// TwinCAT 3 PLC project HrlRbgPlc
// ProgramVersion: 3.1.4026.25
// libraries:
//   NodeTree, * (sulemanali5760)
//   Tc2_MC2, * (Beckhoff Automation GmbH)
//   Tc3_JsonXml, * (Beckhoff Automation GmbH)
//   Tc2_TcpIp, * (Beckhoff Automation GmbH)
//   Tc2_Standard, * (Beckhoff Automation GmbH)
//   Tc2_System, * (Beckhoff Automation GmbH)
//   TcUnit, * (www.tcunit.org)
// project tree:
//   / PlcTask.TcTTO
//   Rack/ GVL_Rack.TcGVL, ST_Slot.TcDUT, ST_SlotAddr.TcDUT, FB_Rack.TcPOU
//   Devices/ E_IPointResult.TcDUT, E_ZoneState.TcDUT, E_AxisKind.TcDUT, I_Axis.TcIO, FB_AxisNc.TcPOU, FB_Axis.TcPOU, FB_ConveyorZone.TcPOU, FB_IPoint.TcPOU
//   Performance/ ST_SrmKinematics.TcDUT, F_DoubleCycleTime.TcPOU, F_LoadHandlingTime.TcPOU, F_MoveTime.TcPOU, F_TravelTime.TcPOU
//   Units/ FB_Srm.TcPOU, E_JogAxis.TcDUT
//   Mfr/ GVL_Mfr.TcGVL, ST_Telegram.TcDUT, FB_MfrInterface.TcPOU, E_MfrLink.TcDUT, ST_TelegramLayout.TcDUT, I_MfrLink.TcIO, FB_TelegramCodec.TcPOU, FB_MfrLinkTcp.TcPOU
//   Machine/ FB_Hrl.TcPOU, FB_MfrEmulator.TcPOU, MAIN.TcPOU
//   Test/ GVL_Test.TcGVL, FB_Axis_Test.TcPOU, FB_ConveyorZone_Test.TcPOU, FB_IPoint_Test.TcPOU, FB_MfrInterface_Test.TcPOU, FB_Rack_Test.TcPOU, FB_Srm_Test.TcPOU, FB_TravelTime_Test.TcPOU, FB_AxisNc_Test.TcPOU, FB_HrlConfig_Test.TcPOU, FB_MfrLinkFake.TcPOU, FB_TelegramCodec_Test.TcPOU, FB_Operation_Test.TcPOU, FB_SafetyInterface_Test.TcPOU, PRG_TEST.TcPOU
//   Config/ ST_RackConfig.TcDUT, ST_AxisConfig.TcDUT, ST_ZoneConfig.TcDUT, ST_HrlConfig.TcDUT, FB_HrlConfig.TcPOU
//   Commissioning/ FB_TeachIn.TcPOU
//   Diag/ E_Fault.TcDUT, FB_Diag.TcPOU
//   Safety/ ST_SafetyStatus.TcDUT, FB_SafetyInterface.TcPOU
//   Hmi/ ST_HmiStatus.TcDUT, ST_HmiCommand.TcDUT, GVL_Hmi.TcGVL, FB_HmiBridge.TcPOU
// real-time tasks:
//   TASK PlcTask: cycle T#10ms, priority 20, ADS port 350
// motion (NC):
//   TASK NC-Task 1 SAF: cycle T#2ms, priority 4, ADS port 501
//   TASK NC-Task 1 SVB: cycle T#10ms, priority 8, ADS port 511
//   AXIS Travel (id 1)
//     Velo: Fast=3000, Maximum=3500
//     OtherSettings: AllowMotionCmdToSlave=true
//     encoder EncType=1
//     drive DrvType=5
//       Analog: VeloReferenz=3500, TorqueSetpointScale=10, ScaleFactorActTorque=0.1
//       TimeComp: TaskDelayCycles=1
//     controller CtrType=1
//       CtrPara: PriorControlFactor=1
//         Observer: BandWidth=20
//   AXIS Hoist (id 2)
//     OtherSettings: AllowMotionCmdToSlave=true
//     encoder EncType=1
//     drive DrvType=5
//       Analog: TorqueSetpointScale=10, ScaleFactorActTorque=0.1
//       TimeComp: TaskDelayCycles=1
//     controller CtrType=1
//       CtrPara: PriorControlFactor=1
//         Observer: BandWidth=20
//   AXIS Fork (id 3)
//     OtherSettings: AllowMotionCmdToSlave=true
//     encoder EncType=1
//     drive DrvType=5
//       Analog: TorqueSetpointScale=10, ScaleFactorActTorque=0.1
//       TimeComp: TaskDelayCycles=1
//     controller CtrType=1
//       CtrPara: PriorControlFactor=1
//         Observer: BandWidth=20
//   AXIS TestAxis (id 4)
//     OtherSettings: AllowMotionCmdToSlave=true
//     encoder EncType=1
//     drive DrvType=5
//       Analog: TorqueSetpointScale=10, ScaleFactorActTorque=0.1
//       TimeComp: TaskDelayCycles=1
//     controller CtrType=1
//       CtrPara: PriorControlFactor=1
//         Observer: BandWidth=20
//   AXIS TestTravel (id 5)
//     Velo: Fast=3000, Maximum=3500
//     OtherSettings: AllowMotionCmdToSlave=true
//     encoder EncType=1
//     drive DrvType=5
//       Analog: VeloReferenz=3500, TorqueSetpointScale=10, ScaleFactorActTorque=0.1
//       TimeComp: TaskDelayCycles=1
//     controller CtrType=1
//       CtrPara: PriorControlFactor=1
//         Observer: BandWidth=20
//   AXIS TestHoist (id 6)
//     OtherSettings: AllowMotionCmdToSlave=true
//     encoder EncType=1
//     drive DrvType=5
//       Analog: TorqueSetpointScale=10, ScaleFactorActTorque=0.1
//       TimeComp: TaskDelayCycles=1
//     controller CtrType=1
//       CtrPara: PriorControlFactor=1
//         Observer: BandWidth=20
//   AXIS TestFork (id 7)
//     OtherSettings: AllowMotionCmdToSlave=true
//     encoder EncType=1
//     drive DrvType=5
//       Analog: TorqueSetpointScale=10, ScaleFactorActTorque=0.1
//       TimeComp: TaskDelayCycles=1
//     controller CtrType=1
//       CtrPara: PriorControlFactor=1
//         Observer: BandWidth=20
// variable links:
//   HrlRbgPlc/HrlRbgPlc Instance <-> NC-Task 1 SAF/Axes/Fork
//     PlcTask Inputs/MAIN.fbPlant.fbSrm.fbForkNc.stAxis.NcToPlc <-> Outputs/ToPlc
//     PlcTask Outputs/MAIN.fbPlant.fbSrm.fbForkNc.stAxis.PlcToNc <-> Inputs/FromPlc
//   HrlRbgPlc/HrlRbgPlc Instance <-> NC-Task 1 SAF/Axes/Hoist
//     PlcTask Inputs/MAIN.fbPlant.fbSrm.fbHoistNc.stAxis.NcToPlc <-> Outputs/ToPlc
//     PlcTask Outputs/MAIN.fbPlant.fbSrm.fbHoistNc.stAxis.PlcToNc <-> Inputs/FromPlc
//   HrlRbgPlc/HrlRbgPlc Instance <-> NC-Task 1 SAF/Axes/TestAxis
//     PlcTask Inputs/PRG_TEST.fbAxisNcTest.fbAxis.stAxis.NcToPlc <-> Outputs/ToPlc
//     PlcTask Outputs/PRG_TEST.fbAxisNcTest.fbAxis.stAxis.PlcToNc <-> Inputs/FromPlc
//   HrlRbgPlc/HrlRbgPlc Instance <-> NC-Task 1 SAF/Axes/TestFork
//     PlcTask Inputs/PRG_TEST.fbAxisNcTest.fbSrmNc.fbForkNc.stAxis.NcToPlc <-> Outputs/ToPlc
//     PlcTask Outputs/PRG_TEST.fbAxisNcTest.fbSrmNc.fbForkNc.stAxis.PlcToNc <-> Inputs/FromPlc
//   HrlRbgPlc/HrlRbgPlc Instance <-> NC-Task 1 SAF/Axes/TestHoist
//     PlcTask Inputs/PRG_TEST.fbAxisNcTest.fbSrmNc.fbHoistNc.stAxis.NcToPlc <-> Outputs/ToPlc
//     PlcTask Outputs/PRG_TEST.fbAxisNcTest.fbSrmNc.fbHoistNc.stAxis.PlcToNc <-> Inputs/FromPlc
//   HrlRbgPlc/HrlRbgPlc Instance <-> NC-Task 1 SAF/Axes/TestTravel
//     PlcTask Inputs/PRG_TEST.fbAxisNcTest.fbSrmNc.fbTravelNc.stAxis.NcToPlc <-> Outputs/ToPlc
//     PlcTask Outputs/PRG_TEST.fbAxisNcTest.fbSrmNc.fbTravelNc.stAxis.PlcToNc <-> Inputs/FromPlc
//   HrlRbgPlc/HrlRbgPlc Instance <-> NC-Task 1 SAF/Axes/Travel
//     PlcTask Inputs/MAIN.fbPlant.fbSrm.fbTravelNc.stAxis.NcToPlc <-> Outputs/ToPlc
//     PlcTask Outputs/MAIN.fbPlant.fbSrm.fbTravelNc.stAxis.PlcToNc <-> Inputs/FromPlc

CONFIGURATION HrlRbgPlc
    RESOURCE PLC ON TwinCAT3
        TASK PlcTask(INTERVAL := T#10ms, PRIORITY := 20);
        PROGRAM MAIN WITH PlcTask : MAIN;
        PROGRAM PRG_TEST WITH PlcTask : PRG_TEST;
    END_RESOURCE
END_CONFIGURATION

// ---- Rack/ST_Slot.TcDUT
TYPE ST_Slot :
STRUCT
    bOccupied : BOOL;
    sLeId     : STRING(20);   // load unit id (pallet barcode)
    bTaught   : BOOL;         // TRUE once the place was measured in teach mode
    lrTaughtX : LREAL;        // measured travel position [m]
    lrTaughtY : LREAL;        // measured hoist position [m]
END_STRUCT
END_TYPE

// ---- Rack/ST_SlotAddr.TcDUT
// Address of a storage place, as the material flow computer sends it.
// Column 0 / level 1 / side 1 is the transfer station (Uebergabeplatz) at the
// front of the aisle, where the pre-zone hands pallets to the RBG.
TYPE ST_SlotAddr :
STRUCT
    nSide   : INT;   // 1 = left, 2 = right (seen from the transfer station)
    nColumn : INT;   // 1..GVL_Rack.cColumns, 0 = transfer station
    nLevel  : INT;   // 1..GVL_Rack.cLevels
END_STRUCT
END_TYPE

// ---- Devices/E_IPointResult.TcDUT
{attribute 'qualified_only'}
{attribute 'strict'}
TYPE E_IPointResult :
(
    eOk         := 0,   // contour fine, barcode read -> may be stored
    eNioContour := 1,   // overhang or too high -> back to the operator
    eNioNoRead  := 2    // barcode not readable -> back to the operator
) DINT;
END_TYPE

// ---- Devices/E_ZoneState.TcDUT
{attribute 'qualified_only'}
{attribute 'strict'}
TYPE E_ZoneState :
(
    eEmpty      := 0,
    eReceiving  := 1,   // motor on, pallet running in
    eOccupied   := 2,   // pallet at the end light barrier, motor off
    eDelivering := 3,   // motor on, pallet running out to the next zone
    eFault      := 4    // jam (light barrier not reached in time) or drive fault
) DINT;
END_TYPE

// ---- Devices/E_AxisKind.TcDUT
// Which implementation drives the RBG axes. Switched in the configuration,
// never in the code: the sequence only talks to I_Axis.
{attribute 'qualified_only'}
{attribute 'strict'}
TYPE E_AxisKind :
(
    eSim := 0,   // FB_Axis: simulated trapezoid profile, simulated time (tests, demo)
    eNc  := 1    // FB_AxisNc: Beckhoff NC axis via Tc2_MC2 (real drive or NC simulation axis)
) INT;
END_TYPE

// ---- Performance/ST_SrmKinematics.TcDUT
TYPE ST_SrmKinematics :
STRUCT
    lrVeloX  : LREAL;   // travel
    lrAccelX : LREAL;
    lrVeloY  : LREAL;   // hoist
    lrAccelY : LREAL;
    lrVeloZ  : LREAL;   // telescopic fork
    lrAccelZ : LREAL;
END_STRUCT
END_TYPE

// ---- Mfr/ST_Telegram.TcDUT
// One telegram between the material flow computer (MFR, e.g. WAMAS) and the PLC.
// The real WAMAS layout is project-specific; this is a typical fixed layout.
TYPE ST_Telegram :
STRUCT
    sType    : STRING(4);    // TORD order, TACK acknowledge, TDON done, TERR error
    nSeq     : UINT;         // sequence number of the sender, +1 per telegram
    nOrder   : DINT;         // transport order number
    sLeId    : STRING(20);   // load unit id
    stSource : ST_SlotAddr;
    stTarget : ST_SlotAddr;
    nStatus  : INT;          // GVL_Mfr status codes, 0 = OK
END_STRUCT
END_TYPE

// ---- Config/ST_RackConfig.TcDUT
// Rack geometry of one aisle. Defaults = the practice plant (GVL_Rack).
// Sizes may not exceed GVL_Rack.cMaxSides / cMaxColumns / cMaxLevels.
TYPE ST_RackConfig :
STRUCT
    nSides          : INT   := GVL_Rack.cSides;
    nColumns        : INT   := GVL_Rack.cColumns;
    nLevels         : INT   := GVL_Rack.cLevels;
    lrPitchX        : LREAL := GVL_Rack.cPitchX;          // column pitch incl. upright [m]
    lrPitchY        : LREAL := GVL_Rack.cPitchY;          // level pitch [m]
    lrOffsetX       : LREAL := GVL_Rack.cOffsetX;         // transfer station -> centre of column 1 [m]
    lrOffsetY       : LREAL := GVL_Rack.cOffsetY;         // fork height at level 1 / station [m]
    lrForkStroke    : LREAL := GVL_Rack.cForkStroke;      // [m]
    lrLiftStroke    : LREAL := GVL_Rack.cLiftStroke;      // [m]
    lrTeachTolerance: LREAL := GVL_Rack.cTeachTolerance;  // [m]
END_STRUCT
END_TYPE

// ---- Config/ST_AxisConfig.TcDUT
TYPE ST_AxisConfig :
STRUCT
    lrVelocity : LREAL := 1.0;   // [m/s]
    lrAccel    : LREAL := 0.5;   // acceleration = deceleration [m/s2]
END_STRUCT
END_TYPE

// ---- Config/ST_ZoneConfig.TcDUT
// Parameters of one conveyor zone (the standard block FB_ConveyorZone).
TYPE ST_ZoneConfig :
STRUCT
    lrLength     : LREAL := 1.6;    // up to the end light barrier [m]
    lrSpeed      : LREAL := 0.2;    // [m/s]
    lrJamTimeout : LREAL := 20.0;   // [s]
    bSimulate    : BOOL  := TRUE;   // FALSE: end light barrier from the real input
END_STRUCT
END_TYPE

// ---- Config/ST_HrlConfig.TcDUT
// Everything an integrator sets per plant. Loaded from HrlConfig.json by
// FB_HrlConfig; every default here is the practice plant, so a missing file
// or a missing entry still gives a working demo.
TYPE ST_HrlConfig :
STRUCT
    stRack    : ST_RackConfig;
    eAxisKind : E_AxisKind := E_AxisKind.eSim;
    stTravel  : ST_AxisConfig := (lrVelocity := 3.0, lrAccel := 0.6);
    stHoist   : ST_AxisConfig := (lrVelocity := 1.5, lrAccel := 0.8);
    stFork    : ST_AxisConfig := (lrVelocity := 0.6, lrAccel := 0.6);
    stInfeed  : ST_ZoneConfig;
    stOutfeed : ST_ZoneConfig := (lrLength := 2.4, lrSpeed := 0.2, lrJamTimeout := 20.0, bSimulate := TRUE);
    lrAckTimeout : LREAL := 5.0;   // MFR must acknowledge TDON within this [s]
    eMfrLink     : E_MfrLink := E_MfrLink.eEmulator;
    nMfrPort     : UINT := 2000;    // TCP port the PLC listens on (eTcp)
    stLayout     : ST_TelegramLayout;
    bSafetySimulate : BOOL := TRUE;   // bench without safety controller (never on a real machine)
END_STRUCT
END_TYPE

// ---- Mfr/E_MfrLink.TcDUT
// Where the transport orders come from.
{attribute 'qualified_only'}
{attribute 'strict'}
TYPE E_MfrLink :
(
    eEmulator := 0,   // FB_MfrEmulator in the PLC (commissioning, demo, tests)
    eTcp      := 1    // real material flow computer over TCP/IP (PLC is the server)
) INT;
END_TYPE

// ---- Mfr/ST_TelegramLayout.TcDUT
// Field widths of the fixed-length ASCII telegram. The field order is fixed:
//   type | seq | order | load unit | source side,column,level | target side,column,level | status
// Numbers are right-aligned with leading zeros, the load unit id is
// left-aligned and padded with spaces. The frame is STX + fields + ETX.
// Defaults give a 52-character telegram.
TYPE ST_TelegramLayout :
STRUCT
    nType   : INT := 4;
    nSeq    : INT := 5;
    nOrder  : INT := 8;
    nLeId   : INT := 20;
    nSide   : INT := 1;
    nColumn : INT := 3;
    nLevel  : INT := 2;
    nStatus : INT := 3;
END_STRUCT
END_TYPE

// ---- Units/E_JogAxis.TcDUT
// Axis the operator jogs in manual mode.
{attribute 'qualified_only'}
{attribute 'strict'}
TYPE E_JogAxis :
(
    eTravel := 0,
    eHoist  := 1,
    eFork   := 2
) INT;
END_TYPE

// ---- Diag/E_Fault.TcDUT
// Plant faults reported by FB_Diag (index into its active list).
{attribute 'qualified_only'}
{attribute 'strict'}
TYPE E_Fault :
(
    eSrmAxis      := 1,   // an RBG axis failed during a job
    eInfeedJam    := 2,
    eOutfeedJam   := 3,
    eMfrAck       := 4,   // MFR did not acknowledge TDON in time
    eMfrLinkDown  := 5,   // TCP link configured but no MFR connected
    eConfig       := 6,   // HrlConfig.json rejected, defaults in use
    eTeachRejected:= 7,   // measured place too far from the drawing
    eSafety       := 8    // safety stop or restart lock active
) INT;
END_TYPE

// ---- Safety/ST_SafetyStatus.TcDUT
// Status bits the safety controller (e.g. TwinSAFE logic) gives the standard
// PLC. The standard PLC only reads them: it never switches safety itself.
// Map each bit to the TwinSAFE group output (see docs/safety/README.md).
TYPE ST_SafetyStatus :
STRUCT
    bSafetyRun  : BOOL;   // safety program running, no group error
    bEStopOk    : BOOL;   // all emergency stops released
    bDoorClosed : BOOL;   // aisle access door closed
    bDoorLocked : BOOL;   // aisle access door guard-locked
    bStoOk      : BOOL;   // drives not in Safe Torque Off
END_STRUCT
END_TYPE

// ---- Hmi/ST_HmiStatus.TcDUT
// Everything the HMI shows (PLC -> HMI). Filled by MAIN every cycle.
TYPE ST_HmiStatus :
STRUCT
    nMode          : INT;          // 0 stop, 1 manual, 2 homing, 3 automatic (E_OpMode)
    bSafetyOk      : BOOL;
    lrTravelPos    : LREAL;        // [m]
    lrHoistPos     : LREAL;        // [m]
    lrForkPos      : LREAL;        // [m]
    bBusy          : BOOL;         // RBG job running
    bFault         : BOOL;         // RBG fault, needs reset
    bJogBlocked    : BOOL;         // jog refused: fork not centred
    sLeOnFork      : STRING(20);
    nJobsDone      : DINT;
    nStored        : DINT;         // emulator counters
    nRetrieved     : DINT;
    bMfrConnected  : BOOL;         // TCP link (always FALSE with the emulator)
    nActiveFaults  : INT;
    sFault1        : STRING(80);   // first four active faults, cause - remedy
    sFault2        : STRING(80);
    sFault3        : STRING(80);
    sFault4        : STRING(80);
    bTeachActive   : BOOL;
    nTaught        : INT;
    bTeachRejected : BOOL;
    sConfigError   : STRING(120);
END_STRUCT
END_TYPE

// ---- Hmi/ST_HmiCommand.TcDUT
// Everything the HMI may command (HMI -> PLC). Buttons that trigger an action
// (teach start/confirm, resets) are evaluated on the rising edge in MAIN.
TYPE ST_HmiCommand :
STRUCT
    bModeStop     : BOOL;       // mode buttons: TRUE while pressed (button state symbol)
    bModeManual   : BOOL;
    bModeHoming   : BOOL;
    bModeAuto     : BOOL;
    nJogAxis      : INT;        // 0 travel, 1 hoist, 2 fork
    bJogFwd       : BOOL;       // held while the button is pressed
    bJogBwd       : BOOL;
    nTeachSide    : INT := 1;
    nTeachColumn  : INT := 1;
    nTeachLevel   : INT := 1;
    bTeachStart   : BOOL;
    bTeachConfirm : BOOL;
    bResetFault   : BOOL;       // RBG fault reset
    bSafetyReset  : BOOL;       // safety acknowledge
END_STRUCT
END_TYPE

// ---- Rack/GVL_Rack.TcGVL
{attribute 'qualified_only'}
VAR_GLOBAL CONSTANT
    // Largest rack the PLC reserves memory for. The real size comes from the
    // configuration (ST_RackConfig) and may be anything up to these.
    cMaxSides   : INT   := 2;
    cMaxColumns : INT   := 60;
    cMaxLevels  : INT   := 16;
    // Defaults = the practice plant: one aisle, single-deep, both sides.
    cSides      : INT   := 2;
    cColumns    : INT   := 20;
    cLevels     : INT   := 8;
    cPitchX     : LREAL := 1.40;   // column pitch incl. upright [m]
    cPitchY     : LREAL := 1.30;   // level pitch [m]
    cOffsetX    : LREAL := 2.00;   // transfer station -> centre of column 1 [m]
    cOffsetY    : LREAL := 0.50;   // fork height at level 1 / transfer station [m]
    cForkStroke : LREAL := 1.10;   // telescopic fork travel into a place [m]
    cLiftStroke : LREAL := 0.10;   // lift to take a pallet off its beams [m]
    // Teach-in: a measured place may differ from the drawing by this much;
    // more means a bent or wrongly built rack -> reject and check the rack.
    cTeachTolerance : LREAL := 0.020;   // [m]
END_VAR

// ---- Mfr/GVL_Mfr.TcGVL
{attribute 'qualified_only'}
VAR_GLOBAL CONSTANT
    cStatusOk         : INT := 0;
    cSlotOccupied     : INT := 10;   // target place occupied
    cSlotEmpty        : INT := 11;   // source place empty
    cContourNio       : INT := 20;   // pallet failed the I-point
    cAckTimeout       : INT := 30;   // MFR did not acknowledge TDON in time
    cWrongSequence    : INT := 40;   // telegram sequence number out of order
    cDuplicateOrder   : INT := 41;   // order number already active / just done
    cInvalidAddress   : INT := 42;
    cSrmBusy          : INT := 43;
    cLeMismatch       : INT := 44;   // load unit at the source is not the one ordered
    cUnknownTelegram  : INT := 45;
    cSrmFault         : INT := 50;
END_VAR

// ---- Test/GVL_Test.TcGVL
{attribute 'qualified_only'}
VAR_GLOBAL
    // Results of the FEM 9.851 double-cycle test, for the performance protocol.
    lrDoubleCycleCalc     : LREAL;   // calculated [s]
    lrDoubleCycleMeasured : LREAL;   // measured in the simulation [s]
    lrDoubleCyclesPerHour : LREAL;   // 3600 / measured
END_VAR

// ---- Hmi/GVL_Hmi.TcGVL
// The only PLC data the HMI uses. Both structs are mapped automatically into
// the TwinCAT HMI server (attribute TcHmiSymbol.AddSymbol).
{attribute 'qualified_only'}
VAR_GLOBAL
    {attribute 'TcHmiSymbol.AddSymbol'}
    stStatus  : ST_HmiStatus;
    {attribute 'TcHmiSymbol.AddSymbol'}
    stCommand : ST_HmiCommand;
END_VAR

// ---- Devices/I_Axis.TcIO
// I_Axis - what the RBG sequence needs from a positioning axis, whatever
// drives it: the simulated FB_Axis or the NC axis FB_AxisNc. Units are metres.
INTERFACE I_Axis

// Drive to an absolute position: eBusy while moving, eDone in position, eError on a fault.
METHOD MoveAbs : E_CmdResult
VAR_INPUT
    lrPos : LREAL;   // target [m]
END_VAR
END_METHOD

// Acknowledge a fault: the axis stops where it is and waits for a new target.
METHOD Reset
VAR_INPUT
END_VAR
END_METHOD

// Stop now (end of a jog, stop mode). The axis then waits for a new target.
METHOD Halt
VAR_INPUT
END_VAR
END_METHOD

// Actual position [m].
PROPERTY ActPos : LREAL
GET
END_GET
END_PROPERTY

PROPERTY Error : BOOL
GET
END_GET
END_PROPERTY

END_INTERFACE

// ---- Mfr/I_MfrLink.TcIO
// I_MfrLink - transport of telegrams between the PLC and the material flow
// computer. FB_MfrInterface only sees telegrams; how they travel (TCP, a test
// double) is behind this interface.
INTERFACE I_MfrLink

// Next received telegram, TRUE if there was one. A frame that could not be
// decoded comes back with sType = 'BAD'.
METHOD Poll : BOOL
VAR_IN_OUT
    stIn : ST_Telegram;
END_VAR
END_METHOD

// Queue a telegram for the MFR. FALSE if not connected or the queue is full.
METHOD Send : BOOL
VAR_INPUT
    stOut : ST_Telegram;
END_VAR
END_METHOD

PROPERTY Connected : BOOL
GET
END_GET
END_PROPERTY

END_INTERFACE

// ---- Machine/MAIN.TcPOU
// MAIN - builds the plant from HrlConfig.json, runs it in the operating mode
// the HMI asks for (eModeRequest), forced to stop while the safety interface
// does not allow motion. With mfr.link = emulator the MFR emulator drives it.
// Watch fbPlant.fbSrm (positions, jobs), fbPlant.fbRack and fbPlant.fbDiag online.
PROGRAM MAIN
VAR
    fbPlant      : FB_Hrl(ipParent := 0, sNodeName := 'HRL');
    fbOpMode     : FB_OpModeHandler;
    fbEmulator   : FB_MfrEmulator;
    fbConfig     : FB_HrlConfig;   // HrlConfig.json from the boot folder; defaults if absent
    fbHmi        : FB_HmiBridge;   // GVL_Hmi <-> plant
    eModeNow     : E_OpMode;
    bInit        : BOOL := TRUE;
END_VAR

IF bInit THEN
    fbConfig();
    IF NOT fbConfig.bDone THEN
        RETURN;   // the plant starts only with its final configuration
    END_IF
    fbPlant.stConfig     := fbConfig.stConfig;
    fbPlant.sConfigError := fbConfig.sError;
    fbOpMode.SetRoot(fbPlant);
    bInit := FALSE;
END_IF

fbHmi.Run(fbPlant, fbEmulator, GVL_Hmi.stCommand, GVL_Hmi.stStatus, eModeNow);
IF fbPlant.bSafetyOk THEN
    eModeNow := fbHmi.eModeRequest;
ELSE
    eModeNow := E_OpMode.eStop;   // safety first: no motion without the safety OK
END_IF
fbOpMode.Mode := eModeNow;
IF fbPlant.stConfig.eMfrLink = E_MfrLink.eEmulator THEN
    fbEmulator.Run(fbPlant);   // no real MFR: the emulator sends the orders
END_IF
fbOpMode.Cyclic();

END_PROGRAM

// ---- Machine/FB_Hrl.TcPOU
// FB_Hrl - the whole practice plant as the root mode node: one aisle with one
// RBG, the rack, the pre-zone with I-point and in-feed/out-feed conveyors, and
// the MFR interface.
// Pre-zone flow: in-feed (pallet already checked at the I-point) -> transfer
// station -> RBG stores it. Retrieved pallets are put on the station and leave
// over the out-feed.
FUNCTION_BLOCK FB_Hrl EXTENDS FB_ModeNode
VAR_INPUT
    stConfig : ST_HrlConfig;   // applied once on the first cycle (set it before)
    sConfigError : STRING(120);   // from FB_HrlConfig; shown as a fault
    stSafety     : ST_SafetyStatus;   // map from the safety controller (TwinSAFE group outputs)
    bSafetyReset : BOOL;              // acknowledge button
    bDoorRequest : BOOL;              // operator wants to enter the aisle
END_VAR
VAR
    fbRack    : FB_Rack;
    fbSrm     : FB_Srm(ipParent := THIS^, sNodeName := 'RBG01');
    fbInfeed  : FB_ConveyorZone(ipParent := THIS^, sNodeName := 'Infeed');
    fbOutfeed : FB_ConveyorZone(ipParent := THIS^, sNodeName := 'Outfeed');
    fbIPoint  : FB_IPoint;
    fbMfr     : FB_MfrInterface;
    fbMfrTcp  : FB_MfrLinkTcp;     // used when stConfig.eMfrLink = eTcp
    fbTeach   : FB_TeachIn;        // guided teach-in (manual mode)
    fbDiag    : FB_Diag;           // active faults for the HMI + TwinCAT logger
    fbSafety  : FB_SafetyInterface;
    bInitDone : BOOL;
    nInStep   : INT;
    sMovingLe : STRING(20);
END_VAR
VAR_OUTPUT
    bStationOutbound : BOOL;   // pallet on the station is leaving (retrieved), not arriving
    bStationReserved : BOOL;   // station held free for a retrieval: the in-feed must wait
    bSafetyOk        : BOOL;   // drives may run; FALSE -> MAIN forces stop mode
    bDoorUnlockReq   : BOOL;   // to the safety controller
END_VAR

METHOD PROTECTED OnCyclic
VAR_INPUT
END_VAR
IF NOT bInitDone THEN
    // The plant is built from the configuration; the code below never changes per site.
    fbRack.stCfg      := stConfig.stRack;
    fbSrm.eAxisKind   := stConfig.eAxisKind;
    fbSrm.stTravelCfg := stConfig.stTravel;
    fbSrm.stHoistCfg  := stConfig.stHoist;
    fbSrm.stForkCfg   := stConfig.stFork;
    ApplyZone(fbInfeed, stConfig.stInfeed);    // same standard block, other parameters
    ApplyZone(fbOutfeed, stConfig.stOutfeed);
    fbMfr.lrAckTimeout := stConfig.lrAckTimeout;
    fbSrm.Init(fbRack);
    fbMfr.Init(fbRack, fbSrm);
    fbTeach.Init(fbRack, fbSrm);
    fbMfrTcp.nPort    := stConfig.nMfrPort;
    fbMfrTcp.stLayout := stConfig.stLayout;
    bInitDone := TRUE;
END_IF
IF stConfig.eMfrLink = E_MfrLink.eTcp THEN
    fbMfrTcp.Cyclic();          // the link stays up in every operating mode
    fbMfr.Serve(fbMfrTcp);
END_IF
fbSafety(stStatus := stSafety, bSimulate := stConfig.bSafetySimulate, bReset := bSafetyReset,
         bDoorRequest := bDoorRequest, bStandstill := NOT fbSrm.bBusy AND NOT fbSrm.bGotoActive);
bSafetyOk      := fbSafety.bDriveEnable;
bDoorUnlockReq := fbSafety.bDoorUnlockReq;
SUPER^.OnCyclic();
fbDiag.Check(E_Fault.eSafety, NOT bSafetyOk, 'Safety stop - check e-stop and aisle door, then acknowledge');
fbDiag.Check(E_Fault.eSrmAxis, fbSrm.bFault, 'RBG axis fault - check the drive, then ResetFault');
fbDiag.Check(E_Fault.eInfeedJam, fbInfeed.eState = E_ZoneState.eFault, 'In-feed jam - clear the pallet, reset the zone');
fbDiag.Check(E_Fault.eOutfeedJam, fbOutfeed.eState = E_ZoneState.eFault, 'Out-feed jam - clear the pallet, reset the zone');
fbDiag.Check(E_Fault.eMfrAck, fbMfr.bAckTimeout, 'MFR did not acknowledge TDON - check the MFR');
fbDiag.Check(E_Fault.eMfrLinkDown, stConfig.eMfrLink = E_MfrLink.eTcp AND NOT fbMfrTcp.bConnected,
             'No MFR connected - check network / MFR port');
fbDiag.Check(E_Fault.eConfig, sConfigError <> '', 'HrlConfig.json rejected - defaults in use, see sConfigError');
fbDiag.Check(E_Fault.eTeachRejected, fbTeach.bLastRejected, 'Teach-in refused - place too far from drawing, check rack');
END_METHOD

METHOD PROTECTED RunAutomatic
VAR_INPUT
END_VAR
VAR
    stStation : ST_SlotAddr := (nSide := 1, nColumn := 0, nLevel := 1);
END_VAR
fbMfr.Cyclic();

// In-feed -> transfer station
CASE nInStep OF
    0:  IF fbInfeed.eState = E_ZoneState.eOccupied AND NOT fbRack.IsOccupied(stStation)
           AND NOT bStationOutbound AND NOT bStationReserved THEN
            sMovingLe := fbInfeed.sLeId;
            nInStep   := 1;
        END_IF
    // Done once our pallet has left the zone. The previous zone may hand over
    // the next pallet in the same cycle, so "zone empty" alone can be missed.
    1:  IF fbInfeed.Deliver() = E_CmdResult.eDone OR fbInfeed.sLeId <> sMovingLe THEN
            fbRack.Put(stStation, sMovingLe);
            nInStep := 0;
        END_IF
END_CASE

// Transfer station -> out-feed (only pallets the RBG brought out)
IF bStationOutbound AND fbRack.IsOccupied(stStation)
   AND fbOutfeed.eState = E_ZoneState.eEmpty THEN
    fbOutfeed.Accept(fbRack.Take(stStation));
    bStationOutbound := FALSE;
    bStationReserved := FALSE;   // station free for the in-feed again
END_IF
IF fbOutfeed.eState = E_ZoneState.eOccupied THEN
    fbOutfeed.Deliver();   // goods-out takes it away
END_IF
END_METHOD

// Called when a retrieval to the station is ordered: that pallet leaves.
METHOD PUBLIC MarkStationOutbound
VAR_INPUT
END_VAR
bStationOutbound := TRUE;
END_METHOD

// Hold the transfer station free for the next retrieval. Without this the
// in-feed refills the station every time the RBG picks a pallet from it, and
// a retrieval never finds the station empty.
METHOD PUBLIC ReserveStation
VAR_INPUT
END_VAR
bStationReserved := TRUE;
END_METHOD

// Manual jog request from the HMI (acts in manual mode only).
METHOD PUBLIC Jog
VAR_INPUT
    eAxis : E_JogAxis;
    bFwd  : BOOL;
    bBwd  : BOOL;
END_VAR
fbSrm.eJogAxis := eAxis;
fbSrm.bJogFwd  := bFwd;
fbSrm.bJogBwd  := bBwd;
END_METHOD

METHOD PRIVATE ApplyZone
VAR_IN_OUT
    fbZone : FB_ConveyorZone;
END_VAR
VAR_INPUT
    stCfg : ST_ZoneConfig;
END_VAR
fbZone.lrLength     := stCfg.lrLength;
fbZone.lrSpeed      := stCfg.lrSpeed;
fbZone.lrJamTimeout := stCfg.lrJamTimeout;
fbZone.bSimulate    := stCfg.bSimulate;
END_METHOD

END_FUNCTION_BLOCK

// ---- Rack/FB_Rack.TcPOU
// FB_Rack - the PLC's picture of the rack: which place is occupied by which
// load unit, and where each place really is (nominal from the drawing, or the
// value measured during teach-in). It is data, not a machine node, so the RBG,
// the MFR interface and the tests all share one instance by reference.
FUNCTION_BLOCK FB_Rack
VAR_INPUT
    stCfg : ST_RackConfig;   // geometry; set once before the first job (FB_Hrl does it from the config)
END_VAR
VAR
    aSlot     : ARRAY[1..GVL_Rack.cMaxSides, 1..GVL_Rack.cMaxColumns, 1..GVL_Rack.cMaxLevels] OF ST_Slot;
    stStation : ST_Slot;   // the transfer station in front of the aisle
END_VAR

METHOD PUBLIC IsStation : BOOL
VAR_INPUT
    stAddr : ST_SlotAddr;
END_VAR
IsStation := stAddr.nColumn = 0 AND stAddr.nLevel = 1 AND stAddr.nSide = 1;
END_METHOD

METHOD PUBLIC IsValid : BOOL
VAR_INPUT
    stAddr : ST_SlotAddr;
END_VAR
IsValid := IsStation(stAddr)
        OR (stAddr.nSide >= 1 AND stAddr.nSide <= stCfg.nSides
            AND stAddr.nColumn >= 1 AND stAddr.nColumn <= stCfg.nColumns
            AND stAddr.nLevel >= 1 AND stAddr.nLevel <= stCfg.nLevels);
END_METHOD

// Pointer to the place record, or 0 for an invalid address.
METHOD PRIVATE Slot : POINTER TO ST_Slot
VAR_INPUT
    stAddr : ST_SlotAddr;
END_VAR
IF IsStation(stAddr) THEN
    Slot := ADR(stStation);
ELSIF IsValid(stAddr) THEN
    Slot := ADR(aSlot[stAddr.nSide, stAddr.nColumn, stAddr.nLevel]);
ELSE
    Slot := 0;
END_IF
END_METHOD

// Travel position of a place from the drawing [m].
METHOD PUBLIC NominalX : LREAL
VAR_INPUT
    stAddr : ST_SlotAddr;
END_VAR
IF IsStation(stAddr) THEN
    NominalX := 0.0;
ELSE
    NominalX := stCfg.lrOffsetX + INT_TO_LREAL(stAddr.nColumn - 1) * stCfg.lrPitchX;
END_IF
END_METHOD

// Hoist position of a place from the drawing [m].
METHOD PUBLIC NominalY : LREAL
VAR_INPUT
    stAddr : ST_SlotAddr;
END_VAR
NominalY := stCfg.lrOffsetY + INT_TO_LREAL(stAddr.nLevel - 1) * stCfg.lrPitchY;
END_METHOD

// Where the RBG drives to: the taught position if there is one, else nominal.
METHOD PUBLIC TargetX : LREAL
VAR_INPUT
    stAddr : ST_SlotAddr;
END_VAR
VAR
    pSlot : POINTER TO ST_Slot;
END_VAR
pSlot := Slot(stAddr);
IF pSlot <> 0 AND_THEN pSlot^.bTaught THEN
    TargetX := pSlot^.lrTaughtX;
ELSE
    TargetX := NominalX(stAddr);
END_IF
END_METHOD

METHOD PUBLIC TargetY : LREAL
VAR_INPUT
    stAddr : ST_SlotAddr;
END_VAR
VAR
    pSlot : POINTER TO ST_Slot;
END_VAR
pSlot := Slot(stAddr);
IF pSlot <> 0 AND_THEN pSlot^.bTaught THEN
    TargetY := pSlot^.lrTaughtY;
ELSE
    TargetY := NominalY(stAddr);
END_IF
END_METHOD

// Store the measured position of a place (teach-in). Returns FALSE and keeps
// the old value if the measurement is further than cTeachTolerance from the
// drawing - that is a rack to check, not a value to learn.
METHOD PUBLIC Teach : BOOL
VAR_INPUT
    stAddr : ST_SlotAddr;
    lrX    : LREAL;   // measured travel position [m] (laser distance sensor)
    lrY    : LREAL;   // measured hoist position [m]
END_VAR
VAR
    pSlot : POINTER TO ST_Slot;
END_VAR
pSlot := Slot(stAddr);
IF pSlot = 0 OR IsStation(stAddr)
   OR ABS(lrX - NominalX(stAddr)) > stCfg.lrTeachTolerance
   OR ABS(lrY - NominalY(stAddr)) > stCfg.lrTeachTolerance THEN
    Teach := FALSE;
    RETURN;
END_IF
pSlot^.lrTaughtX := lrX;
pSlot^.lrTaughtY := lrY;
pSlot^.bTaught   := TRUE;
Teach := TRUE;
END_METHOD

METHOD PUBLIC IsOccupied : BOOL
VAR_INPUT
    stAddr : ST_SlotAddr;
END_VAR
VAR
    pSlot : POINTER TO ST_Slot;
END_VAR
pSlot := Slot(stAddr);
IsOccupied := pSlot <> 0 AND_THEN pSlot^.bOccupied;
END_METHOD

METHOD PUBLIC LeIdAt : STRING(20)
VAR_INPUT
    stAddr : ST_SlotAddr;
END_VAR
VAR
    pSlot : POINTER TO ST_Slot;
END_VAR
pSlot := Slot(stAddr);
IF pSlot <> 0 AND_THEN pSlot^.bOccupied THEN
    LeIdAt := pSlot^.sLeId;
ELSE
    LeIdAt := '';
END_IF
END_METHOD

// Book a load unit into a place. FALSE if the place is invalid or occupied.
METHOD PUBLIC Put : BOOL
VAR_INPUT
    stAddr : ST_SlotAddr;
    sLeId  : STRING(20);
END_VAR
VAR
    pSlot : POINTER TO ST_Slot;
END_VAR
pSlot := Slot(stAddr);
IF pSlot = 0 OR_ELSE pSlot^.bOccupied OR sLeId = '' THEN
    Put := FALSE;
    RETURN;
END_IF
pSlot^.bOccupied := TRUE;
pSlot^.sLeId     := sLeId;
Put := TRUE;
END_METHOD

// Book a load unit out of a place; returns its id, or '' if the place was empty.
METHOD PUBLIC Take : STRING(20)
VAR_INPUT
    stAddr : ST_SlotAddr;
END_VAR
VAR
    pSlot : POINTER TO ST_Slot;
END_VAR
pSlot := Slot(stAddr);
IF pSlot = 0 OR_ELSE NOT pSlot^.bOccupied THEN
    Take := '';
    RETURN;
END_IF
Take := pSlot^.sLeId;
pSlot^.bOccupied := FALSE;
pSlot^.sLeId     := '';
END_METHOD

// First free place, filled column by column from the transfer station
// (short travel first). FALSE if the rack is full.
METHOD PUBLIC FindFree : BOOL
VAR_IN_OUT
    stFound : ST_SlotAddr;
END_VAR
VAR
    nCol, nLvl, nSide : INT;
END_VAR
FOR nCol := 1 TO stCfg.nColumns DO
    FOR nLvl := 1 TO stCfg.nLevels DO
        FOR nSide := 1 TO stCfg.nSides DO
            IF NOT aSlot[nSide, nCol, nLvl].bOccupied THEN
                stFound.nSide   := nSide;
                stFound.nColumn := nCol;
                stFound.nLevel  := nLvl;
                FindFree := TRUE;
                RETURN;
            END_IF
        END_FOR
    END_FOR
END_FOR
FindFree := FALSE;
END_METHOD

END_FUNCTION_BLOCK

// ---- Units/FB_Srm.TcPOU
// FB_Srm - the storage and retrieval machine (Regalbediengeraet, RBG) as a
// mode node. Its three axes are child device nodes, so one Cyclic() on the RBG
// runs the sequence first and then lets the axes move in the same scan.
//
// A job moves one load unit from a source place to a target place (either may
// be the transfer station). The sequence is the classic single cycle:
//   travel+hoist to source -> fork out -> lift -> fork in ->
//   travel+hoist to target (loaded, lifted) -> fork out -> lower -> fork in.
// Two jobs back to back (store, then retrieve) make a double cycle.
FUNCTION_BLOCK FB_Srm EXTENDS FB_ModeNode
VAR_INPUT
    eAxisKind : E_AxisKind := E_AxisKind.eSim;   // simulated axes or NC axes
    stTravelCfg : ST_AxisConfig := (lrVelocity := 3.0, lrAccel := 0.6);
    stHoistCfg  : ST_AxisConfig := (lrVelocity := 1.5, lrAccel := 0.8);
    stForkCfg   : ST_AxisConfig := (lrVelocity := 0.6, lrAccel := 0.6);
    // Manual mode (HMI): hold bJogFwd / bJogBwd to move eJogAxis, release to stop.
    eJogAxis : E_JogAxis := E_JogAxis.eTravel;
    bJogFwd  : BOOL;
    bJogBwd  : BOOL;
END_VAR
VAR_OUTPUT
    bBusy         : BOOL;         // a job is running
    bJobDone      : BOOL;         // last job finished; stays TRUE until the next StartJob
    bFault        : BOOL;         // sequence stopped on an axis fault -> ResetFault
    nJobsDone     : DINT;
    lrLastJobTime : LREAL;        // simulated duration of the last job [s]
    sLeOnFork     : STRING(20);   // load unit currently on the fork
    bJogBlocked   : BOOL;         // jog refused: fork not centred for travel / hoist
    bGotoActive   : BOOL;         // manual: driving to a GotoXY target (teach-in)
END_VAR
VAR
    fbTravel : FB_Axis(ipParent := THIS^, sNodeName := 'Travel');
    fbHoist  : FB_Axis(ipParent := THIS^, sNodeName := 'Hoist');
    fbFork   : FB_Axis(ipParent := THIS^, sNodeName := 'Fork');
    fbTravelNc : FB_AxisNc(ipParent := THIS^, sNodeName := 'TravelNc');
    fbHoistNc  : FB_AxisNc(ipParent := THIS^, sNodeName := 'HoistNc');
    fbForkNc   : FB_AxisNc(ipParent := THIS^, sNodeName := 'ForkNc');
    ipTravel : I_Axis;   // the axes the sequence uses, chosen by eAxisKind
    ipHoist  : I_Axis;
    ipFork   : I_Axis;
    fbCycle  : FB_CycleManager;
    refRack  : REFERENCE TO FB_Rack;
    stSource : ST_SlotAddr;
    stTarget : ST_SlotAddr;
    bJobPending : BOOL;
    lrJobTime   : LREAL;
    lrGotoX     : LREAL;
    lrGotoY     : LREAL;
    bJogging    : BOOL;
END_VAR

// Give the RBG the rack it works on (once, before the first job).
METHOD PUBLIC Init
VAR_INPUT
    fbRackRef : REFERENCE TO FB_Rack;
END_VAR
refRack REF= fbRackRef;
END_METHOD

// Accept a transport job. FALSE if busy, faulted, the addresses are invalid,
// the source is empty or the target is occupied.
METHOD PUBLIC StartJob : BOOL
VAR_INPUT
    stFrom : ST_SlotAddr;
    stTo   : ST_SlotAddr;
END_VAR
StartJob := FALSE;
IF NOT __ISVALIDREF(refRack) OR bJobPending OR bFault THEN
    RETURN;
END_IF
IF NOT refRack.IsValid(stFrom) OR NOT refRack.IsValid(stTo)
   OR NOT refRack.IsOccupied(stFrom) OR refRack.IsOccupied(stTo) THEN
    RETURN;
END_IF
stSource    := stFrom;
stTarget    := stTo;
lrJobTime   := 0.0;
bJobDone    := FALSE;
bJobPending := TRUE;
fbCycle.Reset();   // so the next Call() sees a fresh start edge
StartJob := TRUE;
END_METHOD

// Acknowledge a fault. A load unit still on the fork stays booked on the fork.
METHOD PUBLIC ResetFault
VAR_INPUT
END_VAR
SelectAxes();
ipTravel.Reset();
ipHoist.Reset();
ipFork.Reset();
fbCycle.Reset();
bFault      := FALSE;
bJobPending := FALSE;
END_METHOD

// Travel and hoist together; done when both are in position.
METHOD PRIVATE MoveXY : E_CmdResult
VAR_INPUT
    lrX : LREAL;
    lrY : LREAL;
END_VAR
VAR
    eX, eY : E_CmdResult;
END_VAR
eX := ipTravel.MoveAbs(lrX);
eY := ipHoist.MoveAbs(lrY);
IF eX = E_CmdResult.eError OR eY = E_CmdResult.eError THEN
    MoveXY := E_CmdResult.eError;
ELSIF eX = E_CmdResult.eDone AND eY = E_CmdResult.eDone THEN
    MoveXY := E_CmdResult.eDone;
ELSE
    MoveXY := E_CmdResult.eBusy;
END_IF
END_METHOD

// Fork end position for a place: left side (and the station) negative, right positive.
METHOD PRIVATE ForkPos : LREAL
VAR_INPUT
    stAddr : ST_SlotAddr;
END_VAR
IF stAddr.nSide = 2 THEN
    ForkPos := refRack.stCfg.lrForkStroke;
ELSE
    ForkPos := -refRack.stCfg.lrForkStroke;
END_IF
END_METHOD

METHOD PROTECTED OnCyclic
VAR_INPUT
END_VAR
SelectAxes();
// Axis data from the configuration (defaults = the practice RBG).
fbTravel.lrVelocity   := stTravelCfg.lrVelocity;  fbTravel.lrAccel   := stTravelCfg.lrAccel;
fbHoist.lrVelocity    := stHoistCfg.lrVelocity;   fbHoist.lrAccel    := stHoistCfg.lrAccel;
fbFork.lrVelocity     := stForkCfg.lrVelocity;    fbFork.lrAccel     := stForkCfg.lrAccel;
fbTravelNc.lrVelocity := stTravelCfg.lrVelocity;  fbTravelNc.lrAccel := stTravelCfg.lrAccel;
fbHoistNc.lrVelocity  := stHoistCfg.lrVelocity;   fbHoistNc.lrAccel  := stHoistCfg.lrAccel;
fbForkNc.lrVelocity   := stForkCfg.lrVelocity;    fbForkNc.lrAccel   := stForkCfg.lrAccel;
IF bJobPending THEN
    lrJobTime := lrJobTime + fbTravel.lrCycleTime;
END_IF
SUPER^.OnCyclic();   // dispatch to RunAutomatic / RunManual / ...
bBusy := bJobPending;
END_METHOD

METHOD PROTECTED RunAutomatic
VAR_INPUT
END_VAR
IF NOT __ISVALIDREF(refRack) THEN
    RETURN;
END_IF

fbCycle.Call(bExecute := bJobPending);
CASE fbCycle.Step OF
    0:  fbCycle.Await(MoveXY(refRack.TargetX(stSource), refRack.TargetY(stSource)));
    1:  fbCycle.Await(ipFork.MoveAbs(ForkPos(stSource)));
    2:  IF fbCycle.Await(ipHoist.MoveAbs(refRack.TargetY(stSource) + refRack.stCfg.lrLiftStroke)) THEN
            sLeOnFork := refRack.Take(stSource);   // pallet is now on the fork
        END_IF
    3:  fbCycle.Await(ipFork.MoveAbs(0.0));
    4:  fbCycle.Await(MoveXY(refRack.TargetX(stTarget), refRack.TargetY(stTarget) + refRack.stCfg.lrLiftStroke));
    5:  fbCycle.Await(ipFork.MoveAbs(ForkPos(stTarget)));
    6:  IF fbCycle.Await(ipHoist.MoveAbs(refRack.TargetY(stTarget))) THEN
            refRack.Put(stTarget, sLeOnFork);      // pallet is on the beams
            sLeOnFork := '';
        END_IF
    7:  IF fbCycle.Await(ipFork.MoveAbs(0.0)) THEN
            bJobPending   := FALSE;
            bJobDone      := TRUE;
            nJobsDone     := nJobsDone + 1;
            lrLastJobTime := lrJobTime;
        END_IF
END_CASE

IF fbCycle.Error THEN
    bFault := TRUE;
END_IF
END_METHOD

// Go to the transfer station: fork in first, then travel and hoist.
METHOD PROTECTED RunHoming
VAR_INPUT
END_VAR
IF NOT __ISVALIDREF(refRack) THEN
    RETURN;
END_IF
IF ipFork.MoveAbs(0.0) = E_CmdResult.eDone THEN
    MoveXY(0.0, refRack.stCfg.lrOffsetY);
END_IF
END_METHOD

PROPERTY PUBLIC TravelPos : LREAL
GET
SelectAxes();
TravelPos := ipTravel.ActPos;
END_GET
END_PROPERTY

PROPERTY PUBLIC HoistPos : LREAL
GET
SelectAxes();
HoistPos := ipHoist.ActPos;
END_GET
END_PROPERTY

PROPERTY PUBLIC ForkActPos : LREAL
GET
SelectAxes();
ForkActPos := ipFork.ActPos;
END_GET
END_PROPERTY

// Test and commissioning aid: simulate a fault of the travel drive.
METHOD PUBLIC InjectTravelFault
VAR_INPUT
    bFaultOn : BOOL;
END_VAR
fbTravel.bDriveFault := bFaultOn;
END_METHOD

// Manual mode: drive travel and hoist to a position (fork stays centred).
// Used by teach-in to go to the nominal position of a place.
METHOD PUBLIC GotoXY : BOOL
VAR_INPUT
    lrX : LREAL;
    lrY : LREAL;
END_VAR
IF bFault OR bJobPending THEN
    RETURN;
END_IF
lrGotoX     := lrX;
lrGotoY     := lrY;
bGotoActive := TRUE;
GotoXY      := TRUE;
END_METHOD

// Jog one axis while a button is held; travel and hoist only with the fork
// centred (a fork in the rack would hit the uprights). A GotoXY target has
// priority over jogging.
METHOD PROTECTED RunManual
VAR_INPUT
END_VAR
VAR
    ipAx    : I_Axis;
    lrLimit : LREAL;
END_VAR
IF NOT __ISVALIDREF(refRack) THEN
    RETURN;
END_IF
IF bGotoActive THEN
    IF ABS(ipFork.ActPos) > 0.005 THEN
        ipFork.MoveAbs(0.0);
    ELSIF MoveXY(lrGotoX, lrGotoY) <> E_CmdResult.eBusy THEN
        bGotoActive := FALSE;
    END_IF
    RETURN;
END_IF
CASE eJogAxis OF
    E_JogAxis.eTravel:
        ipAx := ipTravel;
        IF bJogFwd THEN
            lrLimit := refRack.stCfg.lrOffsetX + INT_TO_LREAL(refRack.stCfg.nColumns - 1) * refRack.stCfg.lrPitchX;
        ELSE
            lrLimit := 0.0;
        END_IF
    E_JogAxis.eHoist:
        ipAx := ipHoist;
        IF bJogFwd THEN
            lrLimit := refRack.stCfg.lrOffsetY + INT_TO_LREAL(refRack.stCfg.nLevels - 1) * refRack.stCfg.lrPitchY
                       + refRack.stCfg.lrLiftStroke;
        ELSE
            lrLimit := refRack.stCfg.lrOffsetY;
        END_IF
    E_JogAxis.eFork:
        ipAx := ipFork;
        IF bJogFwd THEN
            lrLimit := refRack.stCfg.lrForkStroke;
        ELSE
            lrLimit := -refRack.stCfg.lrForkStroke;
        END_IF
END_CASE
bJogBlocked := eJogAxis <> E_JogAxis.eFork AND ABS(ipFork.ActPos) > 0.005 AND (bJogFwd OR bJogBwd);
IF (bJogFwd XOR bJogBwd) AND NOT bJogBlocked THEN
    ipAx.MoveAbs(lrLimit);   // runs towards the soft limit while held
    bJogging := TRUE;
ELSIF bJogging THEN
    ipAx.Halt();
    bJogging := FALSE;
END_IF
END_METHOD

// Stop mode: every axis halts. A running job stays pending and the sequence
// resumes from its current step when the mode is set back to automatic.
METHOD PROTECTED RunStop
VAR_INPUT
END_VAR
ipTravel.Halt();
ipHoist.Halt();
ipFork.Halt();
bGotoActive := FALSE;
bJogging    := FALSE;
END_METHOD

// Point the sequence at the simulated or the NC axes. Only the chosen NC
// axes are enabled, so an unlinked NC axis never raises errors in simulation.
METHOD PRIVATE SelectAxes
VAR_INPUT
END_VAR
fbTravelNc.bEnable := eAxisKind = E_AxisKind.eNc;
fbHoistNc.bEnable  := fbTravelNc.bEnable;
fbForkNc.bEnable   := fbTravelNc.bEnable;
IF fbTravelNc.bEnable THEN
    ipTravel := fbTravelNc;
    ipHoist  := fbHoistNc;
    ipFork   := fbForkNc;
ELSE
    ipTravel := fbTravel;
    ipHoist  := fbHoist;
    ipFork   := fbFork;
END_IF
END_METHOD

END_FUNCTION_BLOCK

// ---- Devices/FB_Axis.TcPOU
// FB_Axis - one positioning axis of the RBG (travel, hoist or telescopic fork)
// as a device node. The outside sees one command, MoveAbs(), returning an
// E_CmdResult - same contract as the cylinder in the pick-and-place demo.
//
// There is no drive on a soft-PLC, so the axis simulates itself: a trapezoid
// velocity profile with limited speed and acceleration, integrated once per
// call with lrCycleTime. lrActPos stands for the laser distance sensor value.
// Simulated time (not wall clock) keeps the tests fast and repeatable.
FUNCTION_BLOCK FB_Axis EXTENDS FB_CyclicNode IMPLEMENTS I_Axis
VAR_INPUT
    lrVelocity    : LREAL := 1.0;     // max. speed [m/s]
    lrAccel       : LREAL := 0.5;     // acceleration = deceleration [m/s2]
    lrTolerance   : LREAL := 0.002;   // in-position window [m]
    lrCycleTime   : LREAL := 0.01;    // simulated seconds per call (= PlcTask 10 ms)
    lrMoveTimeout : LREAL := 60.0;    // simulated seconds before a move counts as failed
    bDriveFault   : BOOL;             // drive reports a fault (from the drive / a test)
END_VAR
VAR_OUTPUT
    lrActPos    : LREAL;              // actual position [m] (laser distance sensor)
    lrActVelo   : LREAL;              // actual velocity [m/s]
    bInPosition : BOOL := TRUE;
    bError      : BOOL;
END_VAR
VAR
    lrTarget   : LREAL;
    lrMoveTime : LREAL;
END_VAR

// Drive to an absolute position. eBusy while moving, eDone in position,
// eError on a drive fault or a move that does not arrive in lrMoveTimeout.
METHOD PUBLIC MoveAbs : E_CmdResult
VAR_INPUT
    lrPos : LREAL;   // target [m]
END_VAR
IF ABS(lrPos - lrTarget) > 1.0E-9 THEN   // a new target is a new move
    lrTarget    := lrPos;
    lrMoveTime  := 0.0;
    bInPosition := ABS(lrActPos - lrTarget) <= lrTolerance;
END_IF
IF bError THEN
    MoveAbs := E_CmdResult.eError;
ELSIF bInPosition THEN
    MoveAbs := E_CmdResult.eDone;
ELSE
    MoveAbs := E_CmdResult.eBusy;
END_IF
END_METHOD

// Acknowledge a fault: the axis stops where it is and waits for a new target.
METHOD PUBLIC Reset
VAR_INPUT
END_VAR
bError      := FALSE;
lrActVelo   := 0.0;
lrTarget    := lrActPos;
lrMoveTime  := 0.0;
bInPosition := TRUE;
END_METHOD

METHOD PROTECTED OnCyclic
VAR_INPUT
END_VAR
VAR
    lrDist : LREAL;
    lrDir  : LREAL;
    lrVmax : LREAL;
    lrStep : LREAL;
END_VAR
IF bDriveFault THEN
    lrActVelo := 0.0;
    IF NOT bInPosition THEN
        bError := TRUE;   // a fault while moving fails the move
    END_IF
    RETURN;
END_IF
IF bInPosition OR bError THEN
    lrActVelo := 0.0;
    RETURN;
END_IF

lrDist := lrTarget - lrActPos;
IF lrDist >= 0.0 THEN
    lrDir := 1.0;
ELSE
    lrDir := -1.0;
END_IF

// Fastest speed from which the axis can still stop at the target, measured
// from where it will be after this cycle - braking from the current position
// starts one cycle late and lets the axis arrive faster than physics allows.
lrVmax := MIN(lrVelocity, SQRT(2.0 * lrAccel * MAX(ABS(lrDist) - ABS(lrActVelo) * lrCycleTime, 0.0)));
IF lrActVelo < lrDir * lrVmax THEN
    lrActVelo := MIN(lrActVelo + lrAccel * lrCycleTime, lrDir * lrVmax);
ELSE
    lrActVelo := MAX(lrActVelo - lrAccel * lrCycleTime, lrDir * lrVmax);
END_IF

lrStep := lrActVelo * lrCycleTime;
IF ABS(lrDist - lrStep) <= lrTolerance * 0.5 OR lrDir * (lrDist - lrStep) < 0.0 THEN
    lrActPos    := lrTarget;   // arrived (or would overshoot): snap and stop
    lrActVelo   := 0.0;
    bInPosition := TRUE;
ELSE
    lrActPos := lrActPos + lrStep;
END_IF

lrMoveTime := lrMoveTime + lrCycleTime;
IF NOT bInPosition AND lrMoveTime > lrMoveTimeout THEN
    bError    := TRUE;
    lrActVelo := 0.0;
END_IF
END_METHOD

// Simulated stop: the axis stands where it is (no braking ramp in the simulation).
METHOD PUBLIC Halt
VAR_INPUT
END_VAR
lrActVelo   := 0.0;
lrTarget    := lrActPos;
lrMoveTime  := 0.0;
bInPosition := TRUE;
END_METHOD

PROPERTY PUBLIC ActPos : LREAL
GET
ActPos := lrActPos;
END_GET
END_PROPERTY

PROPERTY PUBLIC Error : BOOL
GET
Error := bError;
END_GET
END_PROPERTY

END_FUNCTION_BLOCK

// ---- Devices/FB_AxisNc.TcPOU
// FB_AxisNc - one RBG axis on a Beckhoff NC axis (Tc2_MC2), with the same
// MoveAbs/Reset contract as the simulated FB_Axis. Link stAxis to an NC axis
// in the System Manager; with no drive linked the NC axis simulates itself, so
// the same code runs on the bench and on the machine.
//
// The PLC works in metres, the NC axis in its own unit (default mm):
// lrScale converts (1000 = NC unit mm).
FUNCTION_BLOCK FB_AxisNc EXTENDS FB_CyclicNode IMPLEMENTS I_Axis
VAR_INPUT
    bEnable     : BOOL;              // FALSE: block does nothing (axis not used)
    lrVelocity  : LREAL := 1.0;      // [m/s]
    lrAccel     : LREAL := 0.5;      // acceleration = deceleration [m/s2]
    lrTolerance : LREAL := 0.002;    // in-position window [m]
    lrScale     : LREAL := 1000.0;   // NC units per metre
END_VAR
VAR_OUTPUT
    lrActPos    : LREAL;             // actual position [m]
    lrActVelo   : LREAL;             // actual velocity [m/s]
    bInPosition : BOOL;
    bError      : BOOL;
    nErrorId    : UDINT;             // NC error code (Beckhoff NC error list)
END_VAR
VAR
    stAxis     : AXIS_REF;           // link to the NC axis
    fbPower    : MC_Power;
    fbReset    : MC_Reset;
    fbMove     : MC_MoveAbsolute;
    fbHalt     : MC_Halt;
    bHaltReq   : BOOL;
    lrTarget   : LREAL;
    bHasTarget : BOOL;
    nMoveStep  : INT;                // 0 idle, 1 new target (Execute low), 2 moving
    bResetReq  : BOOL;
END_VAR

METHOD PUBLIC MoveAbs : E_CmdResult
VAR_INPUT
    lrPos : LREAL;   // target [m]
END_VAR
IF NOT bHasTarget OR ABS(lrPos - lrTarget) > 1.0E-9 THEN   // a new target is a new move
    lrTarget    := lrPos;
    bHasTarget  := TRUE;
    nMoveStep   := 1;
    bInPosition := FALSE;
END_IF
IF bError THEN
    MoveAbs := E_CmdResult.eError;
ELSIF bInPosition THEN
    MoveAbs := E_CmdResult.eDone;
ELSE
    MoveAbs := E_CmdResult.eBusy;
END_IF
END_METHOD

METHOD PUBLIC Reset
VAR_INPUT
END_VAR
bError     := FALSE;
nErrorId   := 0;
bResetReq  := TRUE;
bHasTarget := FALSE;
nMoveStep  := 0;
END_METHOD

// Stop with the configured deceleration (MC_Halt); then wait for a new target.
METHOD PUBLIC Halt
VAR_INPUT
END_VAR
IF nMoveStep <> 0 OR NOT bInPosition THEN
    bHaltReq := TRUE;
END_IF
nMoveStep   := 0;
bHasTarget  := FALSE;
bInPosition := TRUE;
fbMove(Axis := stAxis, Execute := FALSE);
END_METHOD

METHOD PROTECTED OnCyclic
VAR_INPUT
END_VAR
IF NOT bEnable THEN
    RETURN;
END_IF
stAxis.ReadStatus();
lrActPos  := stAxis.NcToPlc.ActPos / lrScale;
lrActVelo := stAxis.NcToPlc.ActVelo / lrScale;

fbReset(Axis := stAxis, Execute := bResetReq);
IF fbReset.Done OR fbReset.Error THEN
    bResetReq := FALSE;
    fbReset(Axis := stAxis, Execute := FALSE);
END_IF
fbPower(Axis := stAxis, Enable := NOT bResetReq, Enable_Positive := TRUE,
        Enable_Negative := TRUE, Override := 100.0);

fbHalt(Axis := stAxis, Execute := bHaltReq, Deceleration := lrAccel * lrScale, Jerk := 0.0);
IF bHaltReq AND (fbHalt.Done OR fbHalt.Error) THEN
    bHaltReq := FALSE;
    fbHalt(Axis := stAxis, Execute := FALSE);
END_IF

// Execute needs a rising edge per target: one cycle low, then high until done.
CASE nMoveStep OF
    1:  fbMove(Axis := stAxis, Execute := FALSE);
        IF fbPower.Status AND NOT bResetReq THEN
            nMoveStep := 2;
        END_IF
    2:  fbMove(Axis := stAxis, Execute := TRUE, Position := lrTarget * lrScale,
               Velocity := lrVelocity * lrScale, Acceleration := lrAccel * lrScale,
               Deceleration := lrAccel * lrScale, Jerk := 0.0);
        IF fbMove.Done THEN
            nMoveStep   := 0;
            bInPosition := TRUE;   // the NC's own position window decides "done"
            fbMove(Axis := stAxis, Execute := FALSE);
        END_IF
END_CASE

IF fbMove.Error OR fbPower.Error OR stAxis.Status.Error THEN
    bError    := TRUE;
    nMoveStep := 0;
    IF stAxis.Status.Error THEN
        nErrorId := stAxis.Status.ErrorID;
    ELSIF fbMove.Error THEN
        nErrorId := fbMove.ErrorID;
    ELSE
        nErrorId := fbPower.ErrorID;
    END_IF
    fbMove(Axis := stAxis, Execute := FALSE);
END_IF
END_METHOD

PROPERTY PUBLIC ActPos : LREAL
GET
ActPos := lrActPos;
END_GET
END_PROPERTY

PROPERTY PUBLIC Error : BOOL
GET
Error := bError;
END_GET
END_PROPERTY

END_FUNCTION_BLOCK

// ---- Devices/FB_ConveyorZone.TcPOU
// FB_ConveyorZone - one roller or chain conveyor zone for pallets, as a
// standard block: every zone of the pre-zone is an instance of this FB and the
// zones differ only in their parameters (length, speed, jam timeout). That is
// the "Parametrierung" of a standard library on site.
//
// A zone holds at most one pallet. Accept() starts receiving, the end light
// barrier stops it (eOccupied), Deliver() runs it out until the light barrier
// is free again. A transport that takes longer than lrJamTimeout is a jam.
// bSimulate fakes the end light barrier from the pallet position.
FUNCTION_BLOCK FB_ConveyorZone EXTENDS FB_CyclicNode
VAR_INPUT
    lrLength       : LREAL := 1.6;    // zone length up to the end light barrier [m]
    lrSpeed        : LREAL := 0.2;    // conveyor speed [m/s]
    lrPalletLength : LREAL := 1.2;    // pallet length in transport direction [m]
    lrJamTimeout   : LREAL := 20.0;   // simulated seconds per transport before a jam
    lrCycleTime    : LREAL := 0.01;
    bSimulate      : BOOL := TRUE;
    bEndSensor     : BOOL;            // end light barrier (map to the terminal)
    bDriveFault    : BOOL;
END_VAR
VAR_OUTPUT
    bMotorOn : BOOL;                  // map to the motor contactor / roller drive
    eState   : E_ZoneState;
    sLeId    : STRING(20);            // pallet currently in the zone
END_VAR
VAR
    lrPallet    : LREAL;              // simulated position of the pallet front [m]
    lrStateTime : LREAL;
END_VAR

// Take over a pallet from the previous zone. Only an empty zone accepts.
METHOD PUBLIC Accept : BOOL
VAR_INPUT
    sId : STRING(20);
END_VAR
IF eState <> E_ZoneState.eEmpty OR sId = '' THEN
    Accept := FALSE;
    RETURN;
END_IF
sLeId       := sId;
lrPallet    := 0.0;
lrStateTime := 0.0;
eState      := E_ZoneState.eReceiving;
Accept      := TRUE;
END_METHOD

// Run the pallet out. eBusy until the zone is empty again (= eDone),
// eError on a fault. An empty zone has nothing to deliver and reports eDone.
METHOD PUBLIC Deliver : E_CmdResult
VAR_INPUT
END_VAR
IF eState = E_ZoneState.eOccupied THEN
    eState      := E_ZoneState.eDelivering;
    lrStateTime := 0.0;
END_IF
CASE eState OF
    E_ZoneState.eEmpty:  Deliver := E_CmdResult.eDone;
    E_ZoneState.eFault:  Deliver := E_CmdResult.eError;
ELSE
    Deliver := E_CmdResult.eBusy;
END_CASE
END_METHOD

// After clearing a jam on site: the zone is empty again.
METHOD PUBLIC Reset
VAR_INPUT
END_VAR
eState      := E_ZoneState.eEmpty;
sLeId       := '';
lrPallet    := 0.0;
lrStateTime := 0.0;
bMotorOn    := FALSE;
END_METHOD

METHOD PROTECTED OnCyclic
VAR_INPUT
END_VAR
bMotorOn := eState = E_ZoneState.eReceiving OR eState = E_ZoneState.eDelivering;

IF bMotorOn THEN
    IF bDriveFault THEN
        eState := E_ZoneState.eFault;
    ELSE
        lrStateTime := lrStateTime + lrCycleTime;
        IF lrStateTime > lrJamTimeout THEN
            eState := E_ZoneState.eFault;   // light barrier not reached / not freed in time
        END_IF
    END_IF
END_IF

IF bSimulate THEN
    IF eState = E_ZoneState.eReceiving OR eState = E_ZoneState.eDelivering THEN
        lrPallet := lrPallet + lrSpeed * lrCycleTime;
    END_IF
    bEndSensor := eState <> E_ZoneState.eEmpty AND eState <> E_ZoneState.eFault
                  AND lrPallet >= lrLength AND lrPallet < lrLength + lrPalletLength;
END_IF

CASE eState OF
    E_ZoneState.eReceiving:
        IF bEndSensor THEN
            eState := E_ZoneState.eOccupied;
        END_IF
    E_ZoneState.eDelivering:
        IF NOT bEndSensor THEN
            eState := E_ZoneState.eEmpty;   // pallet has left the zone
            sLeId  := '';
        END_IF
END_CASE

bMotorOn := eState = E_ZoneState.eReceiving OR eState = E_ZoneState.eDelivering;
END_METHOD

END_FUNCTION_BLOCK

// ---- Devices/FB_IPoint.TcPOU
// FB_IPoint - identification point (I-Punkt) in front of the warehouse: the
// contour check light barriers and the barcode reader decide whether a pallet
// may go into the rack. Every pallet that is stored has passed this check.
FUNCTION_BLOCK FB_IPoint
VAR_INPUT
    bOverhangFront : BOOL;   // light barriers: TRUE = goods stick out
    bOverhangBack  : BOOL;
    bOverhangLeft  : BOOL;
    bOverhangRight : BOOL;
    bTooHigh       : BOOL;
    sBarcode       : STRING(20);   // empty = no read
END_VAR
VAR_OUTPUT
    nChecked : DINT;
    nNio     : DINT;
END_VAR

METHOD PUBLIC Check : E_IPointResult
VAR_INPUT
END_VAR
nChecked := nChecked + 1;
IF bOverhangFront OR bOverhangBack OR bOverhangLeft OR bOverhangRight OR bTooHigh THEN
    Check := E_IPointResult.eNioContour;
ELSIF sBarcode = '' THEN
    Check := E_IPointResult.eNioNoRead;
ELSE
    Check := E_IPointResult.eOk;
END_IF
IF Check <> E_IPointResult.eOk THEN
    nNio := nNio + 1;
END_IF
END_METHOD

END_FUNCTION_BLOCK

// ---- Mfr/FB_MfrInterface.TcPOU
// FB_MfrInterface - the PLC side of the telegram interface to the material
// flow computer. Every incoming telegram is checked before anything moves:
// sequence number, duplicate order, valid addresses, RBG free, source really
// occupied by the ordered load unit, target free. The answer is TACK (accepted)
// or TERR with a status code. When the RBG finishes, the interface sends TDON
// and expects the MFR to acknowledge it within lrAckTimeout.
FUNCTION_BLOCK FB_MfrInterface
VAR_INPUT
    lrCycleTime  : LREAL := 0.01;
    lrAckTimeout : LREAL := 5.0;   // simulated seconds for the MFR to acknowledge TDON
END_VAR
VAR_OUTPUT
    stOutbox     : ST_Telegram;    // last unsolicited telegram (TDON / TERR) for the MFR
    nOutboxCount : DINT;           // +1 per new outbox telegram (edge for the sender)
    nLastStatus  : INT;
    bAckTimeout  : BOOL;
END_VAR
VAR
    refRack      : REFERENCE TO FB_Rack;
    refSrm       : REFERENCE TO FB_Srm;
    nExpectedSeq : UINT := 1;
    nSendSeq     : UINT;
    nActiveOrder : DINT;
    nLastOrder   : DINT;
    bAwaitAck    : BOOL;
    lrAckWait    : LREAL;
    nOutboxSent  : DINT;   // outbox telegrams already handed to the link
END_VAR

METHOD PUBLIC Init
VAR_INPUT
    fbRackRef : REFERENCE TO FB_Rack;
    fbSrmRef  : REFERENCE TO FB_Srm;
END_VAR
refRack REF= fbRackRef;
refSrm  REF= fbSrmRef;
END_METHOD

METHOD PRIVATE Reply : ST_Telegram
VAR_INPUT
    sType   : STRING(4);
    stIn    : ST_Telegram;
    nStatus : INT;
END_VAR
nSendSeq       := nSendSeq + 1;
Reply          := stIn;
Reply.sType    := sType;
Reply.nSeq     := nSendSeq;
Reply.nStatus  := nStatus;
nLastStatus    := nStatus;
END_METHOD

// Handle one telegram from the MFR and return the immediate answer.
METHOD PUBLIC Receive : ST_Telegram
VAR_INPUT
    stIn : ST_Telegram;
END_VAR
IF NOT __ISVALIDREF(refRack) OR NOT __ISVALIDREF(refSrm) THEN
    RETURN;
END_IF

// 1. Sequence: a lost or repeated telegram must never move a pallet.
IF stIn.nSeq <> nExpectedSeq THEN
    Receive := Reply('TERR', stIn, GVL_Mfr.cWrongSequence);
    RETURN;
END_IF
nExpectedSeq := nExpectedSeq + 1;

IF stIn.sType = 'TACK' THEN
    // MFR acknowledges our TDON
    IF bAwaitAck AND stIn.nOrder = nLastOrder THEN
        bAwaitAck := FALSE;
        lrAckWait := 0.0;
    END_IF
    RETURN;   // no answer to an acknowledgement
END_IF

IF stIn.sType <> 'TORD' THEN
    Receive := Reply('TERR', stIn, GVL_Mfr.cUnknownTelegram);
    RETURN;
END_IF

// 2. Transport order: check everything before the RBG moves.
IF stIn.nOrder = nActiveOrder OR stIn.nOrder = nLastOrder THEN
    Receive := Reply('TERR', stIn, GVL_Mfr.cDuplicateOrder);
ELSIF NOT refRack.IsValid(stIn.stSource) OR NOT refRack.IsValid(stIn.stTarget) THEN
    Receive := Reply('TERR', stIn, GVL_Mfr.cInvalidAddress);
ELSIF nActiveOrder <> 0 OR refSrm.bBusy OR refSrm.bFault THEN
    Receive := Reply('TERR', stIn, GVL_Mfr.cSrmBusy);
ELSIF NOT refRack.IsOccupied(stIn.stSource) THEN
    Receive := Reply('TERR', stIn, GVL_Mfr.cSlotEmpty);
ELSIF refRack.IsOccupied(stIn.stTarget) THEN
    Receive := Reply('TERR', stIn, GVL_Mfr.cSlotOccupied);
ELSIF refRack.LeIdAt(stIn.stSource) <> stIn.sLeId THEN
    Receive := Reply('TERR', stIn, GVL_Mfr.cLeMismatch);
ELSIF refSrm.StartJob(stIn.stSource, stIn.stTarget) THEN
    nActiveOrder := stIn.nOrder;
    Receive := Reply('TACK', stIn, GVL_Mfr.cStatusOk);
ELSE
    Receive := Reply('TERR', stIn, GVL_Mfr.cSrmBusy);
END_IF
END_METHOD

// Call every cycle: reports the end of the active order and watches the ack.
METHOD PUBLIC Cyclic
VAR_INPUT
END_VAR
VAR
    stDone : ST_Telegram;
END_VAR
IF NOT __ISVALIDREF(refSrm) THEN
    RETURN;
END_IF

IF nActiveOrder <> 0 THEN
    stDone.nOrder := nActiveOrder;
    IF refSrm.bJobDone THEN
        stOutbox     := Reply('TDON', stDone, GVL_Mfr.cStatusOk);
        nOutboxCount := nOutboxCount + 1;
        nLastOrder   := nActiveOrder;
        nActiveOrder := 0;
        bAwaitAck    := TRUE;
        lrAckWait    := 0.0;
    ELSIF refSrm.bFault THEN
        stOutbox     := Reply('TERR', stDone, GVL_Mfr.cSrmFault);
        nOutboxCount := nOutboxCount + 1;
        nLastOrder   := nActiveOrder;
        nActiveOrder := 0;
    END_IF
END_IF

IF bAwaitAck THEN
    lrAckWait := lrAckWait + lrCycleTime;
    IF lrAckWait > lrAckTimeout THEN
        bAwaitAck   := FALSE;
        bAckTimeout := TRUE;   // shown as a fault; the order itself is done
        nLastStatus := GVL_Mfr.cAckTimeout;
    END_IF
END_IF
END_METHOD

PROPERTY PUBLIC ActiveOrder : DINT
GET
ActiveOrder := nActiveOrder;
END_GET
END_PROPERTY

PROPERTY PUBLIC AwaitingAck : BOOL
GET
AwaitingAck := bAwaitAck;
END_GET
END_PROPERTY

// Call every cycle when the MFR is a real system: takes one telegram from the
// link, runs the same checks as Receive() and sends the answer, then sends any
// new unsolicited telegram (TDON / TERR) from the outbox. An undecodable frame
// is answered with TERR 45 without touching the sequence count.
METHOD PUBLIC Serve
VAR_INPUT
    ipLink : I_MfrLink;
END_VAR
VAR
    stIn    : ST_Telegram;
    stReply : ST_Telegram;
END_VAR
IF ipLink = 0 THEN
    RETURN;
END_IF
IF ipLink.Poll(stIn) THEN
    IF stIn.sType = 'BAD' THEN
        stReply := Reply('TERR', stIn, GVL_Mfr.cUnknownTelegram);
    ELSE
        stReply := Receive(stIn);
    END_IF
    IF stReply.sType <> '' THEN
        ipLink.Send(stReply);
    END_IF
END_IF
IF nOutboxCount <> nOutboxSent AND ipLink.Connected THEN
    IF ipLink.Send(stOutbox) THEN
        nOutboxSent := nOutboxCount;
    END_IF
END_IF
END_METHOD

END_FUNCTION_BLOCK

// ---- Mfr/FB_MfrLinkTcp.TcPOU
// FB_MfrLinkTcp - TCP/IP server for the material flow computer (TF6310,
// Tc2_TcpIp). The PLC listens on nPort; one MFR connects. Every telegram is
// framed as STX (16#02) + fixed-length text + ETX (16#03). Received frames are
// decoded into a small inbox, telegrams to send wait in a small outbox.
// A lost connection closes the socket and waits for the MFR to reconnect.
// Call Cyclic() every PLC cycle.
FUNCTION_BLOCK FB_MfrLinkTcp IMPLEMENTS I_MfrLink
VAR_INPUT
    nPort    : UINT := 2000;
    stLayout : ST_TelegramLayout;
END_VAR
VAR_OUTPUT
    bConnected : BOOL;
    nErrId     : UDINT;   // last socket error (TF6310 error list)
    nBadFrames : UDINT;
END_VAR
VAR
    fbListen : FB_SocketListen;
    fbAccept : FB_SocketAccept;
    fbRecv   : FB_SocketReceive;
    fbSend   : FB_SocketSend;
    fbClose  : FB_SocketClose;
    fbRetry  : TON;
    fbCodec  : FB_TelegramCodec;
    hListener : T_HSOCKET;
    hSocket   : T_HSOCKET;
    nState    : INT;
    aRx       : ARRAY[0..1023] OF BYTE;
    aFrame    : ARRAY[0..255] OF BYTE;   // frame being collected (0-terminated)
    nFrameLen : INT;
    bInFrame  : BOOL;
    aTx       : ARRAY[0..257] OF BYTE;
    bSending  : BOOL;
    aInbox    : ARRAY[0..7] OF ST_Telegram;
    nInHead, nInCount : INT;
    aOutbox   : ARRAY[0..7] OF STRING(255);
    nOutHead, nOutCount : INT;
END_VAR

METHOD PUBLIC Cyclic
VAR_INPUT
END_VAR
VAR
    i : UDINT;
    pFrame : POINTER TO STRING(255);
    stTel  : ST_Telegram;
    sTx    : STRING(255);
END_VAR
fbCodec.stLayout := stLayout;
CASE nState OF
    0:  // open the listening socket
        fbListen(sSrvNetId := '', sLocalHost := '', nLocalPort := nPort, bExecute := TRUE);
        IF NOT fbListen.bBusy THEN
            fbListen(bExecute := FALSE);
            IF fbListen.bError THEN
                nErrId := fbListen.nErrId;
                nState := 90;
            ELSE
                hListener := fbListen.hListener;
                nState := 1;
            END_IF
        END_IF
    1:  // wait for the MFR to connect
        fbAccept(sSrvNetId := '', hListener := hListener, bExecute := TRUE);
        IF NOT fbAccept.bBusy THEN
            fbAccept(bExecute := FALSE);
            IF fbAccept.bError THEN
                nErrId := fbAccept.nErrId;
                nState := 91;
            ELSIF fbAccept.bAccepted THEN
                hSocket    := fbAccept.hSocket;
                bConnected := TRUE;
                bInFrame   := FALSE;
                nState     := 2;
            END_IF
        END_IF
    2:  // connected: receive and send
        fbRecv(sSrvNetId := '', hSocket := hSocket, cbLen := SIZEOF(aRx), pDest := ADR(aRx), bExecute := TRUE);
        IF NOT fbRecv.bBusy THEN
            fbRecv(bExecute := FALSE);
            IF fbRecv.bError THEN
                nErrId := fbRecv.nErrId;
                nState := 80;
            ELSIF fbRecv.nRecBytes > 0 THEN
                FOR i := 0 TO fbRecv.nRecBytes - 1 DO
                    IF aRx[i] = 16#02 THEN            // STX: new frame
                        bInFrame  := TRUE;
                        nFrameLen := 0;
                    ELSIF aRx[i] = 16#03 AND bInFrame THEN   // ETX: frame complete
                        bInFrame := FALSE;
                        aFrame[nFrameLen] := 0;
                        pFrame := ADR(aFrame);
                        IF NOT fbCodec.Decode(pFrame^, stTel) THEN
                            stTel.sType := 'BAD';
                            nBadFrames := nBadFrames + 1;
                        END_IF
                        PushIn(stTel);
                    ELSIF bInFrame AND nFrameLen < 255 THEN
                        aFrame[nFrameLen] := aRx[i];
                        nFrameLen := nFrameLen + 1;
                    END_IF
                END_FOR
            END_IF
        END_IF
        IF bSending THEN
            fbSend(bExecute := TRUE);
            IF NOT fbSend.bBusy THEN
                fbSend(bExecute := FALSE);
                bSending := FALSE;
                IF fbSend.bError THEN
                    nErrId := fbSend.nErrId;
                    nState := 80;
                END_IF
            END_IF
        ELSIF nOutCount > 0 THEN
            sTx := aOutbox[nOutHead];
            nOutHead  := (nOutHead + 1) MOD 8;
            nOutCount := nOutCount - 1;
            aTx[0] := 16#02;
            MEMCPY(destAddr := ADR(aTx[1]), srcAddr := ADR(sTx), n := INT_TO_UDINT(LEN(sTx)));
            aTx[LEN(sTx) + 1] := 16#03;
            fbSend(sSrvNetId := '', hSocket := hSocket, cbLen := INT_TO_UDINT(LEN(sTx) + 2),
                   pSrc := ADR(aTx), bExecute := TRUE);
            bSending := TRUE;
        END_IF
    80: // connection lost: close it and wait for the next one
        fbClose(sSrvNetId := '', hSocket := hSocket, bExecute := TRUE);
        IF NOT fbClose.bBusy THEN
            fbClose(bExecute := FALSE);
            bConnected := FALSE;
            bSending   := FALSE;
            nOutCount  := 0;
            nState     := 1;
        END_IF
    90, 91: // socket error: retry after 2 s (90 = listen again, 91 = accept again)
        fbRetry(IN := TRUE, PT := T#2S);
        IF fbRetry.Q THEN
            fbRetry(IN := FALSE);
            IF nState = 90 THEN
                nState := 0;
            ELSE
                nState := 1;
            END_IF
        END_IF
END_CASE
END_METHOD

METHOD PRIVATE PushIn
VAR_INPUT
    stTel : ST_Telegram;
END_VAR
IF nInCount < 8 THEN   // a full inbox drops the frame; the MFR repeats on timeout
    aInbox[(nInHead + nInCount) MOD 8] := stTel;
    nInCount := nInCount + 1;
END_IF
END_METHOD

METHOD PUBLIC Poll : BOOL
VAR_IN_OUT
    stIn : ST_Telegram;
END_VAR
IF nInCount > 0 THEN
    stIn     := aInbox[nInHead];
    nInHead  := (nInHead + 1) MOD 8;
    nInCount := nInCount - 1;
    Poll     := TRUE;
END_IF
END_METHOD

METHOD PUBLIC Send : BOOL
VAR_INPUT
    stOut : ST_Telegram;
END_VAR
fbCodec.stLayout := stLayout;
IF bConnected AND nOutCount < 8 THEN
    aOutbox[(nOutHead + nOutCount) MOD 8] := fbCodec.Encode(stOut);
    nOutCount := nOutCount + 1;
    Send := TRUE;
END_IF
END_METHOD

PROPERTY PUBLIC Connected : BOOL
GET
Connected := bConnected;
END_GET
END_PROPERTY

END_FUNCTION_BLOCK

// ---- Mfr/FB_TelegramCodec.TcPOU
// FB_TelegramCodec - ST_Telegram <-> fixed-length ASCII text (without STX/ETX).
// The field widths come from stLayout (configuration), the order is fixed (see
// ST_TelegramLayout). Decode refuses a frame of the wrong length or with a
// non-digit in a number field, so a garbled telegram can never move a pallet.
FUNCTION_BLOCK FB_TelegramCodec
VAR_INPUT
    stLayout : ST_TelegramLayout;
END_VAR
VAR
    nPos : INT;   // read position while decoding (1-based, as MID)
END_VAR

METHOD PUBLIC FrameLength : INT
VAR_INPUT
END_VAR
FrameLength := stLayout.nType + stLayout.nSeq + stLayout.nOrder + stLayout.nLeId
             + 2 * (stLayout.nSide + stLayout.nColumn + stLayout.nLevel) + stLayout.nStatus;
END_METHOD

METHOD PUBLIC Encode : STRING(255)
VAR_INPUT
    stTel : ST_Telegram;
END_VAR
VAR
    sAll : STRING(255);   // telegram so far (reading Encode itself would be a recursive call)
    sTmp : STRING(255);   // one field; CONCAT must not take a string function call directly (error 3202)
END_VAR
sAll := Text(stTel.sType, stLayout.nType);
sTmp := Digits(UINT_TO_DINT(stTel.nSeq), stLayout.nSeq);                sAll := CONCAT(sAll, sTmp);
sTmp := Digits(stTel.nOrder, stLayout.nOrder);                          sAll := CONCAT(sAll, sTmp);
sTmp := Text(stTel.sLeId, stLayout.nLeId);                              sAll := CONCAT(sAll, sTmp);
sTmp := Digits(INT_TO_DINT(stTel.stSource.nSide), stLayout.nSide);      sAll := CONCAT(sAll, sTmp);
sTmp := Digits(INT_TO_DINT(stTel.stSource.nColumn), stLayout.nColumn);  sAll := CONCAT(sAll, sTmp);
sTmp := Digits(INT_TO_DINT(stTel.stSource.nLevel), stLayout.nLevel);    sAll := CONCAT(sAll, sTmp);
sTmp := Digits(INT_TO_DINT(stTel.stTarget.nSide), stLayout.nSide);      sAll := CONCAT(sAll, sTmp);
sTmp := Digits(INT_TO_DINT(stTel.stTarget.nColumn), stLayout.nColumn);  sAll := CONCAT(sAll, sTmp);
sTmp := Digits(INT_TO_DINT(stTel.stTarget.nLevel), stLayout.nLevel);    sAll := CONCAT(sAll, sTmp);
sTmp := Digits(INT_TO_DINT(stTel.nStatus), stLayout.nStatus);           sAll := CONCAT(sAll, sTmp);
Encode := sAll;
END_METHOD

// TRUE and stTel filled if sFrame is a well-formed telegram; FALSE otherwise.
METHOD PUBLIC Decode : BOOL
VAR_INPUT
    sFrame : STRING(255);
END_VAR
VAR_IN_OUT
    stTel : ST_Telegram;
END_VAR
VAR
    stNew : ST_Telegram;
    bOk   : BOOL := TRUE;
    sPart : STRING(255);
END_VAR
IF LEN(sFrame) <> FrameLength() THEN
    RETURN;
END_IF
nPos := 1;
sPart                  := Field(sFrame, stLayout.nType);
stNew.sType            := Trimmed(sPart);
sPart := Field(sFrame, stLayout.nSeq);
stNew.nSeq             := DINT_TO_UINT(Number(sPart, bOk));
sPart := Field(sFrame, stLayout.nOrder);
stNew.nOrder           := Number(sPart, bOk);
sPart                  := Field(sFrame, stLayout.nLeId);
stNew.sLeId            := Trimmed(sPart);
sPart := Field(sFrame, stLayout.nSide);
stNew.stSource.nSide   := DINT_TO_INT(Number(sPart, bOk));
sPart := Field(sFrame, stLayout.nColumn);
stNew.stSource.nColumn := DINT_TO_INT(Number(sPart, bOk));
sPart := Field(sFrame, stLayout.nLevel);
stNew.stSource.nLevel  := DINT_TO_INT(Number(sPart, bOk));
sPart := Field(sFrame, stLayout.nSide);
stNew.stTarget.nSide   := DINT_TO_INT(Number(sPart, bOk));
sPart := Field(sFrame, stLayout.nColumn);
stNew.stTarget.nColumn := DINT_TO_INT(Number(sPart, bOk));
sPart := Field(sFrame, stLayout.nLevel);
stNew.stTarget.nLevel  := DINT_TO_INT(Number(sPart, bOk));
sPart := Field(sFrame, stLayout.nStatus);
stNew.nStatus          := DINT_TO_INT(Number(sPart, bOk));
IF bOk THEN
    stTel  := stNew;
    Decode := TRUE;
END_IF
END_METHOD

// Next nWidth characters from nPos on; advances nPos.
METHOD PRIVATE Field : STRING(255)
VAR_INPUT
    sFrame : STRING(255);
    nWidth : INT;
END_VAR
Field := MID(sFrame, nWidth, nPos);
nPos  := nPos + nWidth;
END_METHOD

// Digits-only field to DINT. A non-digit clears bOk.
METHOD PRIVATE Number : DINT
VAR_INPUT
    sField : STRING(255);
END_VAR
VAR_IN_OUT
    bOk : BOOL;
END_VAR
VAR
    i : INT;
    pC : POINTER TO BYTE;
END_VAR
IF LEN(sField) = 0 THEN
    bOk := FALSE;
    RETURN;
END_IF
pC := ADR(sField);
FOR i := 0 TO LEN(sField) - 1 DO
    IF pC[i] < 16#30 OR pC[i] > 16#39 THEN   // '0'..'9'
        bOk := FALSE;
        RETURN;
    END_IF
END_FOR
Number := STRING_TO_DINT(sField);
END_METHOD

// n right-aligned with leading zeros in nWidth characters (keeps the last nWidth digits).
METHOD PRIVATE Digits : STRING(255)
VAR_INPUT
    n      : DINT;
    nWidth : INT;
END_VAR
VAR
    sTmp : STRING(255);
END_VAR
sTmp := DINT_TO_STRING(ABS(n));
WHILE LEN(sTmp) < nWidth DO
    sTmp := CONCAT('0', sTmp);
END_WHILE
Digits := RIGHT(sTmp, nWidth);
END_METHOD

// s left-aligned, padded with spaces / cut to nWidth characters.
METHOD PRIVATE Text : STRING(255)
VAR_INPUT
    sTmp      : STRING(255);
    nWidth : INT;
END_VAR
VAR
    sOut : STRING(255);
END_VAR
sOut := LEFT(sTmp, nWidth);
WHILE LEN(sOut) < nWidth DO
    sOut := CONCAT(sOut, ' ');
END_WHILE
Text := sOut;
END_METHOD

// s without trailing spaces.
METHOD PRIVATE Trimmed : STRING(255)
VAR_INPUT
    sTmp : STRING(255);
END_VAR
VAR
    sOut : STRING(255);
END_VAR
sOut := sTmp;
WHILE LEN(sOut) > 0 AND_THEN RIGHT(sOut, 1) = ' ' DO
    sOut := LEFT(sOut, LEN(sOut) - 1);
END_WHILE
Trimmed := sOut;
END_METHOD

END_FUNCTION_BLOCK

// ---- Commissioning/FB_TeachIn.TcPOU
// FB_TeachIn - guided teach-in of rack places, in manual mode:
//   1. Start(place): the RBG drives to the nominal position from the drawing.
//   2. The operator jogs travel / hoist until the fork lines up with the beams.
//   3. Confirm(): the measured position is stored in the rack, or refused if it
//      is further than the teach tolerance from the drawing (check the rack).
FUNCTION_BLOCK FB_TeachIn
VAR_OUTPUT
    stPlace       : ST_SlotAddr;   // place being taught
    bActive       : BOOL;          // a place is selected
    nTaught       : INT;
    nRejected     : INT;
    bLastRejected : BOOL;
END_VAR
VAR
    refRack : REFERENCE TO FB_Rack;
    refSrm  : REFERENCE TO FB_Srm;
END_VAR

METHOD PUBLIC Init
VAR_INPUT
    fbRackRef : REFERENCE TO FB_Rack;
    fbSrmRef  : REFERENCE TO FB_Srm;
END_VAR
refRack REF= fbRackRef;
refSrm  REF= fbSrmRef;
END_METHOD

// Select a place and drive to its nominal position. FALSE for an invalid
// place, the station, or an RBG that cannot move now.
METHOD PUBLIC Start : BOOL
VAR_INPUT
    stAddr : ST_SlotAddr;
END_VAR
IF NOT __ISVALIDREF(refRack) OR NOT __ISVALIDREF(refSrm) THEN
    RETURN;
END_IF
IF NOT refRack.IsValid(stAddr) OR refRack.IsStation(stAddr) THEN
    RETURN;
END_IF
IF refSrm.GotoXY(refRack.NominalX(stAddr), refRack.NominalY(stAddr)) THEN
    stPlace := stAddr;
    bActive := TRUE;
    Start   := TRUE;
END_IF
END_METHOD

// Store where the RBG stands now as the position of the selected place.
METHOD PUBLIC Confirm : BOOL
VAR_INPUT
END_VAR
IF NOT bActive OR_ELSE refSrm.bGotoActive THEN
    RETURN;   // nothing selected, or still driving there
END_IF
bLastRejected := NOT refRack.Teach(stPlace, refSrm.TravelPos, refSrm.HoistPos);
IF bLastRejected THEN
    nRejected := nRejected + 1;
ELSE
    nTaught := nTaught + 1;
    bActive := FALSE;
    Confirm := TRUE;
END_IF
END_METHOD

END_FUNCTION_BLOCK

// ---- Diag/FB_Diag.TcPOU
// FB_Diag - plant fault list. Call Check() for every fault condition each
// cycle. A fault that becomes active is written once to the TwinCAT logger
// (ADSLOGSTR, visible in the XAE Error List and the logger) with its cause and
// remedy, and stays in aText until the condition clears. The HMI shows aText.
// (Event classes of the TwinCAT EventLogger need the XAE type editor; this
// block uses the logger directly so it builds and runs headless.)
FUNCTION_BLOCK FB_Diag
VAR CONSTANT
    cMaxFault : INT := 16;
END_VAR
VAR_OUTPUT
    nActive : INT;                                // faults active now
    nRaised : UDINT;                              // faults raised since start
    aText   : ARRAY[1..cMaxFault] OF STRING(80);  // '' = not active
END_VAR
VAR
    aActive : ARRAY[1..cMaxFault] OF BOOL;
END_VAR

METHOD PUBLIC Check
VAR_INPUT
    eFault     : E_Fault;
    bCondition : BOOL;
    sText      : STRING(80);   // cause - remedy
END_VAR
VAR
    nIdx : INT;
END_VAR
nIdx := TO_INT(eFault);
IF nIdx < 1 OR nIdx > cMaxFault THEN
    RETURN;
END_IF
IF bCondition AND NOT aActive[nIdx] THEN
    aActive[nIdx] := TRUE;
    aText[nIdx]   := sText;
    nActive := nActive + 1;
    nRaised := nRaised + 1;
    ADSLOGSTR(msgCtrlMask := ADSLOG_MSGTYPE_ERROR OR ADSLOG_MSGTYPE_LOG,
              msgFmtStr := 'HRL fault: %s', strArg := sText);
ELSIF NOT bCondition AND aActive[nIdx] THEN
    aActive[nIdx] := FALSE;
    aText[nIdx]   := '';
    nActive := nActive - 1;
END_IF
END_METHOD

END_FUNCTION_BLOCK

// ---- Safety/FB_SafetyInterface.TcPOU
// FB_SafetyInterface - standard-PLC side of the safety concept. NOT a safety
// function: the safety controller stops the machine on its own; this block
// makes the standard program follow it and adds what the standard side owns:
//   - drive enable and automatic only while every safety bit is OK
//   - restart lock: after any drop, nothing restarts until bReset (rising edge)
//     with all bits OK again (no automatic restart, cf. EN ISO 13849 / EN 528)
//   - door unlock request only while the RBG stands still
// Template only: the integrator validates the whole safety concept per machine.
FUNCTION_BLOCK FB_SafetyInterface
VAR_INPUT
    stStatus      : ST_SafetyStatus;
    bSimulate     : BOOL;   // bench without safety hardware: status counts as OK
    bReset        : BOOL;   // operator acknowledge (rising edge)
    bDoorRequest  : BOOL;   // operator wants to enter the aisle
    bStandstill   : BOOL;   // RBG not moving
END_VAR
VAR_OUTPUT
    bDriveEnable   : BOOL;  // standard enable of the axes / automatic allowed
    bRestartLock   : BOOL;  // a safety bit dropped; waits for bReset
    bDoorUnlockReq : BOOL;  // request to the safety controller to unlock the door
END_VAR
VAR
    fbResetEdge : R_TRIG;
    bAllOk      : BOOL;
    bStarted    : BOOL;
END_VAR

bAllOk := bSimulate OR (stStatus.bSafetyRun AND stStatus.bEStopOk AND stStatus.bDoorClosed
                        AND stStatus.bDoorLocked AND stStatus.bStoOk);
fbResetEdge(CLK := bReset);
IF NOT bStarted THEN            // power-up counts as a drop: acknowledge first
    bRestartLock := NOT bSimulate;
    bStarted     := TRUE;
END_IF
IF NOT bAllOk THEN
    bRestartLock := TRUE;
ELSIF fbResetEdge.Q THEN
    bRestartLock := FALSE;
END_IF
bDriveEnable   := bAllOk AND NOT bRestartLock;
bDoorUnlockReq := bDoorRequest AND bStandstill;

END_FUNCTION_BLOCK

// ---- Machine/FB_MfrEmulator.TcPOU
// FB_MfrEmulator - stands in for the material flow computer (WAMAS) so the
// plant runs on a soft-PLC with nothing connected. It feeds new pallets into
// the in-feed, orders each one into the rack, and after every third store
// orders the oldest pallet back out: stores and retrievals alternate like in
// a real warehouse. It acknowledges every TDON, as the real MFR must.
// Commissioning only - a real plant gets these telegrams from the MFR.
FUNCTION_BLOCK FB_MfrEmulator
VAR_INPUT
    bEnable : BOOL := TRUE;
END_VAR
VAR_OUTPUT
    nStored    : DINT;
    nRetrieved : DINT;
    stLastReply : ST_Telegram;
END_VAR
VAR
    nSeq        : UINT;
    nOrder      : DINT;
    nNextLe     : DINT := 1;
    nSeenOutbox : DINT;
    aStored     : ARRAY[1..400] OF ST_SlotAddr;   // FIFO of stored places
    nHead       : DINT := 1;
    nTail       : DINT := 1;
    nStoresSinceRetrieve : DINT;
    bRetrieving : BOOL;
END_VAR

METHOD PUBLIC Run
VAR_IN_OUT
    fbPlant : FB_Hrl;
END_VAR
VAR
    stTel     : ST_Telegram;
    stStation : ST_SlotAddr := (nSide := 1, nColumn := 0, nLevel := 1);
    stFree    : ST_SlotAddr;
END_VAR
IF NOT bEnable THEN
    RETURN;
END_IF

// Acknowledge every TDON the PLC sends.
IF fbPlant.fbMfr.nOutboxCount <> nSeenOutbox THEN
    nSeenOutbox := fbPlant.fbMfr.nOutboxCount;
    IF fbPlant.fbMfr.stOutbox.sType = 'TDON' THEN
        nSeq := nSeq + 1;
        stTel.sType  := 'TACK';
        stTel.nSeq   := nSeq;
        stTel.nOrder := fbPlant.fbMfr.stOutbox.nOrder;
        fbPlant.fbMfr.Receive(stTel);
        IF bRetrieving THEN
            nRetrieved  := nRetrieved + 1;
            bRetrieving := FALSE;
        END_IF
    END_IF
END_IF

// Feed a new pallet when the in-feed is empty (pallet assumed checked at the I-point).
IF fbPlant.fbInfeed.eState = E_ZoneState.eEmpty THEN
    fbPlant.fbInfeed.Accept(CONCAT('LE', RIGHT(CONCAT('0000', DINT_TO_STRING(nNextLe)), 4)));
    nNextLe := nNextLe + 1;
END_IF

IF fbPlant.fbMfr.ActiveOrder <> 0 OR fbPlant.fbMfr.AwaitingAck OR fbPlant.fbSrm.bBusy THEN
    RETURN;   // one order at a time
END_IF

IF nStoresSinceRetrieve >= 3 AND nTail > nHead AND NOT bRetrieving
   AND NOT fbPlant.fbRack.IsOccupied(stStation) THEN
    // retrieve the oldest pallet to the station
    nSeq   := nSeq + 1;
    nOrder := nOrder + 1;
    stTel.sType    := 'TORD';
    stTel.nSeq     := nSeq;
    stTel.nOrder   := nOrder;
    stTel.stSource := aStored[nHead];
    stTel.stTarget := stStation;
    stTel.sLeId    := fbPlant.fbRack.LeIdAt(aStored[nHead]);
    stLastReply := fbPlant.fbMfr.Receive(stTel);
    IF stLastReply.sType = 'TACK' THEN
        nHead := nHead + 1;
        bRetrieving := TRUE;
        nStoresSinceRetrieve := 0;
        fbPlant.MarkStationOutbound();
    END_IF
ELSIF fbPlant.fbRack.IsOccupied(stStation) AND NOT fbPlant.bStationOutbound
      AND fbPlant.fbRack.FindFree(stFree) AND nTail <= 400 THEN
    // store the pallet waiting on the station
    nSeq   := nSeq + 1;
    nOrder := nOrder + 1;
    stTel.sType    := 'TORD';
    stTel.nSeq     := nSeq;
    stTel.nOrder   := nOrder;
    stTel.stSource := stStation;
    stTel.stTarget := stFree;
    stTel.sLeId    := fbPlant.fbRack.LeIdAt(stStation);
    stLastReply := fbPlant.fbMfr.Receive(stTel);
    IF stLastReply.sType = 'TACK' THEN
        aStored[nTail] := stFree;
        nTail   := nTail + 1;
        nStored := nStored + 1;
        nStoresSinceRetrieve := nStoresSinceRetrieve + 1;
        IF nStoresSinceRetrieve >= 3 THEN
            fbPlant.ReserveStation();   // the next station slot is for a retrieval
        END_IF
    END_IF
END_IF
END_METHOD

END_FUNCTION_BLOCK

// ---- Config/FB_HrlConfig.TcPOU
// FB_HrlConfig - loads the plant configuration once at start-up.
// Call it every cycle until bDone. It reads sFileName from the TwinCAT boot
// folder, parses the JSON and checks every value. A missing file is not an
// error: the plant runs with the built-in defaults (bFileFound = FALSE).
// A file that does not parse or holds a value out of range sets bError and
// sError and also leaves the defaults in place - a bad config never half-applies.
FUNCTION_BLOCK FB_HrlConfig
VAR_INPUT
    sFileName : STRING := 'HrlConfig.json';   // in the boot folder (PATH_BOOTPATH)
END_VAR
VAR_OUTPUT
    bDone      : BOOL;
    bFileFound : BOOL;
    bError     : BOOL;
    sError     : STRING(120);
    stConfig   : ST_HrlConfig;
END_VAR
VAR
    fbOpen  : FB_FileOpen;
    fbRead  : FB_FileRead;
    fbClose : FB_FileClose;
    fbJson  : FB_JsonDomParser;
    hFile   : UINT;
    nStep   : INT;
    bReadOk : BOOL;
    nLen    : UDINT;
    sText   : STRING(8191);
    pEnd    : POINTER TO BYTE;
END_VAR

CASE nStep OF
    0:  fbOpen(sNetId := '', sPathName := sFileName, nMode := FOPEN_MODEREAD OR FOPEN_MODETEXT,
               ePath := PATH_BOOTPATH, bExecute := TRUE);
        nStep := 1;
    1:  fbOpen(bExecute := TRUE);
        IF NOT fbOpen.bBusy THEN
            fbOpen(bExecute := FALSE);
            IF fbOpen.bError THEN       // no file: keep the defaults
                bFileFound := FALSE;
                bDone      := TRUE;
                nStep      := 10;
            ELSE
                hFile := fbOpen.hFile;
                nStep := 2;
            END_IF
        END_IF
    2:  fbRead(sNetId := '', hFile := hFile, pReadBuff := ADR(sText),
               cbReadLen := SIZEOF(sText) - 1, bExecute := TRUE);
        nStep := 3;
    3:  fbRead(bExecute := TRUE);
        IF NOT fbRead.bBusy THEN
            fbRead(bExecute := FALSE);
            bReadOk := NOT fbRead.bError;
            nLen    := fbRead.cbRead;
            nStep   := 4;
        END_IF
    4:  fbClose(sNetId := '', hFile := hFile, bExecute := TRUE);
        nStep := 5;
    5:  fbClose(bExecute := TRUE);
        IF NOT fbClose.bBusy THEN
            fbClose(bExecute := FALSE);
            bFileFound := TRUE;
            IF bReadOk THEN
                pEnd  := ADR(sText) + nLen;   // terminate the string after the bytes read
                pEnd^ := 0;
                Parse(sText);
            ELSE
                bError := TRUE;
                sError := CONCAT('cannot read ', sFileName);
            END_IF
            bDone := TRUE;
            nStep := 10;
        END_IF
END_CASE

// Parse a JSON text into stConfig. Missing entries keep their default.
// FALSE (and stConfig unchanged) if the text is not JSON or a value is out of range.
METHOD PUBLIC Parse : BOOL
VAR_IN_OUT CONSTANT
    sJson : STRING;
END_VAR
VAR
    stNew  : ST_HrlConfig;   // starts as the defaults
    jDoc, jRack, jAxes, jConv, jMfr, jKind, jLayout, jSafety : SJsonValue;
END_VAR
bError := FALSE;
sError := '';
jDoc := fbJson.ParseDocument(sJson);
IF jDoc = 0 THEN
    bError := TRUE;
    sError := 'config is not valid JSON';
    RETURN;
END_IF
jRack := fbJson.FindMember(jDoc, 'rack');
IF jRack <> 0 THEN
    stNew.stRack.nSides           := LREAL_TO_INT(ReadNum(jRack, 'sides', INT_TO_LREAL(stNew.stRack.nSides)));
    stNew.stRack.nColumns         := LREAL_TO_INT(ReadNum(jRack, 'columns', INT_TO_LREAL(stNew.stRack.nColumns)));
    stNew.stRack.nLevels          := LREAL_TO_INT(ReadNum(jRack, 'levels', INT_TO_LREAL(stNew.stRack.nLevels)));
    stNew.stRack.lrPitchX         := ReadNum(jRack, 'pitchX', stNew.stRack.lrPitchX);
    stNew.stRack.lrPitchY         := ReadNum(jRack, 'pitchY', stNew.stRack.lrPitchY);
    stNew.stRack.lrOffsetX        := ReadNum(jRack, 'offsetX', stNew.stRack.lrOffsetX);
    stNew.stRack.lrOffsetY        := ReadNum(jRack, 'offsetY', stNew.stRack.lrOffsetY);
    stNew.stRack.lrForkStroke     := ReadNum(jRack, 'forkStroke', stNew.stRack.lrForkStroke);
    stNew.stRack.lrLiftStroke     := ReadNum(jRack, 'liftStroke', stNew.stRack.lrLiftStroke);
    stNew.stRack.lrTeachTolerance := ReadNum(jRack, 'teachTolerance', stNew.stRack.lrTeachTolerance);
END_IF
jAxes := fbJson.FindMember(jDoc, 'axes');
IF jAxes <> 0 THEN
    jKind := fbJson.FindMember(jAxes, 'kind');
    IF jKind <> 0 THEN
        IF fbJson.GetString(jKind) = 'nc' THEN
            stNew.eAxisKind := E_AxisKind.eNc;
        ELSIF fbJson.GetString(jKind) = 'sim' THEN
            stNew.eAxisKind := E_AxisKind.eSim;
        ELSE
            bError := TRUE;
            sError := 'axes.kind must be sim or nc';
            RETURN;
        END_IF
    END_IF
    stNew.stTravel := ReadAxis(jAxes, 'travel', stNew.stTravel);
    stNew.stHoist  := ReadAxis(jAxes, 'hoist', stNew.stHoist);
    stNew.stFork   := ReadAxis(jAxes, 'fork', stNew.stFork);
END_IF
jConv := fbJson.FindMember(jDoc, 'conveyors');
IF jConv <> 0 THEN
    stNew.stInfeed  := ReadZone(jConv, 'infeed', stNew.stInfeed);
    stNew.stOutfeed := ReadZone(jConv, 'outfeed', stNew.stOutfeed);
END_IF
jMfr := fbJson.FindMember(jDoc, 'mfr');
IF jMfr <> 0 THEN
    stNew.lrAckTimeout := ReadNum(jMfr, 'ackTimeout', stNew.lrAckTimeout);
    stNew.nMfrPort     := LREAL_TO_UINT(ReadNum(jMfr, 'port', UINT_TO_LREAL(stNew.nMfrPort)));
    jKind := fbJson.FindMember(jMfr, 'link');
    IF jKind <> 0 THEN
        IF fbJson.GetString(jKind) = 'tcp' THEN
            stNew.eMfrLink := E_MfrLink.eTcp;
        ELSIF fbJson.GetString(jKind) = 'emulator' THEN
            stNew.eMfrLink := E_MfrLink.eEmulator;
        ELSE
            bError := TRUE;
            sError := 'mfr.link must be emulator or tcp';
            RETURN;
        END_IF
    END_IF
    jLayout := fbJson.FindMember(jMfr, 'layout');
    IF jLayout <> 0 THEN
        stNew.stLayout.nType   := LREAL_TO_INT(ReadNum(jLayout, 'type', INT_TO_LREAL(stNew.stLayout.nType)));
        stNew.stLayout.nSeq    := LREAL_TO_INT(ReadNum(jLayout, 'seq', INT_TO_LREAL(stNew.stLayout.nSeq)));
        stNew.stLayout.nOrder  := LREAL_TO_INT(ReadNum(jLayout, 'order', INT_TO_LREAL(stNew.stLayout.nOrder)));
        stNew.stLayout.nLeId   := LREAL_TO_INT(ReadNum(jLayout, 'leId', INT_TO_LREAL(stNew.stLayout.nLeId)));
        stNew.stLayout.nSide   := LREAL_TO_INT(ReadNum(jLayout, 'side', INT_TO_LREAL(stNew.stLayout.nSide)));
        stNew.stLayout.nColumn := LREAL_TO_INT(ReadNum(jLayout, 'column', INT_TO_LREAL(stNew.stLayout.nColumn)));
        stNew.stLayout.nLevel  := LREAL_TO_INT(ReadNum(jLayout, 'level', INT_TO_LREAL(stNew.stLayout.nLevel)));
        stNew.stLayout.nStatus := LREAL_TO_INT(ReadNum(jLayout, 'status', INT_TO_LREAL(stNew.stLayout.nStatus)));
    END_IF
END_IF
jSafety := fbJson.FindMember(jDoc, 'safety');
IF jSafety <> 0 THEN
    jKind := fbJson.FindMember(jSafety, 'simulate');
    IF jKind <> 0 THEN
        stNew.bSafetySimulate := fbJson.GetBool(jKind);
    END_IF
END_IF
IF NOT Validate(stNew) THEN
    bError := TRUE;
    RETURN;
END_IF
stConfig := stNew;
Parse := TRUE;
END_METHOD

METHOD PRIVATE ReadNum : LREAL
VAR_INPUT
    jParent   : SJsonValue;
    sName     : STRING;
    lrDefault : LREAL;
END_VAR
VAR
    j : SJsonValue;
END_VAR
j := fbJson.FindMember(jParent, sName);
IF j = 0 THEN
    ReadNum := lrDefault;
ELSE
    ReadNum := fbJson.GetDouble(j);
END_IF
END_METHOD

METHOD PRIVATE ReadAxis : ST_AxisConfig
VAR_INPUT
    jParent   : SJsonValue;
    sName     : STRING;
    stDefault : ST_AxisConfig;
END_VAR
VAR
    j : SJsonValue;
END_VAR
ReadAxis := stDefault;
j := fbJson.FindMember(jParent, sName);
IF j <> 0 THEN
    ReadAxis.lrVelocity := ReadNum(j, 'velocity', stDefault.lrVelocity);
    ReadAxis.lrAccel    := ReadNum(j, 'accel', stDefault.lrAccel);
END_IF
END_METHOD

METHOD PRIVATE ReadZone : ST_ZoneConfig
VAR_INPUT
    jParent   : SJsonValue;
    sName     : STRING;
    stDefault : ST_ZoneConfig;
END_VAR
VAR
    j, jSim : SJsonValue;
END_VAR
ReadZone := stDefault;
j := fbJson.FindMember(jParent, sName);
IF j <> 0 THEN
    ReadZone.lrLength     := ReadNum(j, 'length', stDefault.lrLength);
    ReadZone.lrSpeed      := ReadNum(j, 'speed', stDefault.lrSpeed);
    ReadZone.lrJamTimeout := ReadNum(j, 'jamTimeout', stDefault.lrJamTimeout);
    jSim := fbJson.FindMember(j, 'simulate');
    IF jSim <> 0 THEN
        ReadZone.bSimulate := fbJson.GetBool(jSim);
    END_IF
END_IF
END_METHOD

// Range check of a whole configuration; names the first bad value in sError.
METHOD PRIVATE Validate : BOOL
VAR_INPUT
    stChk : ST_HrlConfig;
END_VAR
Validate := FALSE;
IF stChk.stRack.nSides < 1 OR stChk.stRack.nSides > GVL_Rack.cMaxSides THEN
    sError := 'rack.sides out of range';
ELSIF stChk.stRack.nColumns < 1 OR stChk.stRack.nColumns > GVL_Rack.cMaxColumns THEN
    sError := 'rack.columns out of range';
ELSIF stChk.stRack.nLevels < 1 OR stChk.stRack.nLevels > GVL_Rack.cMaxLevels THEN
    sError := 'rack.levels out of range';
ELSIF stChk.stRack.lrPitchX <= 0.0 OR stChk.stRack.lrPitchY <= 0.0 OR stChk.stRack.lrForkStroke <= 0.0
   OR stChk.stRack.lrLiftStroke <= 0.0 OR stChk.stRack.lrTeachTolerance <= 0.0 THEN
    sError := 'rack dimensions must be > 0';
ELSIF NOT AxisOk(stChk.stTravel) OR NOT AxisOk(stChk.stHoist) OR NOT AxisOk(stChk.stFork) THEN
    sError := 'axis velocity / accel must be in 0..10';
ELSIF stChk.stInfeed.lrLength <= 0.0 OR stChk.stInfeed.lrSpeed <= 0.0 OR stChk.stInfeed.lrJamTimeout <= 0.0
   OR stChk.stOutfeed.lrLength <= 0.0 OR stChk.stOutfeed.lrSpeed <= 0.0 OR stChk.stOutfeed.lrJamTimeout <= 0.0 THEN
    sError := 'conveyor length / speed / jamTimeout must be > 0';
ELSIF stChk.lrAckTimeout <= 0.0 THEN
    sError := 'mfr.ackTimeout must be > 0';
ELSIF stChk.nMfrPort = 0 THEN
    sError := 'mfr.port must be 1..65535';
ELSIF stChk.stLayout.nType < 1 OR stChk.stLayout.nType > 4 OR stChk.stLayout.nLeId < 1 OR stChk.stLayout.nLeId > 20
   OR NOT WidthOk(stChk.stLayout.nSeq) OR NOT WidthOk(stChk.stLayout.nOrder) OR NOT WidthOk(stChk.stLayout.nSide)
   OR NOT WidthOk(stChk.stLayout.nColumn) OR NOT WidthOk(stChk.stLayout.nLevel) OR NOT WidthOk(stChk.stLayout.nStatus) THEN
    sError := 'mfr.layout: type 1..4, leId 1..20, numbers 1..9 characters';
ELSE
    Validate := TRUE;
END_IF
END_METHOD

METHOD PRIVATE AxisOk : BOOL
VAR_INPUT
    stChk : ST_AxisConfig;
END_VAR
AxisOk := stChk.lrVelocity > 0.0 AND stChk.lrVelocity <= 10.0 AND stChk.lrAccel > 0.0 AND stChk.lrAccel <= 10.0;
END_METHOD

// A number field fits a DINT with 1..9 digits.
METHOD PRIVATE WidthOk : BOOL
VAR_INPUT
    nWidth : INT;
END_VAR
WidthOk := nWidth >= 1 AND nWidth <= 9;
END_METHOD

END_FUNCTION_BLOCK

// ---- Hmi/FB_HmiBridge.TcPOU
// FB_HmiBridge - copies the plant state into ST_HmiStatus and applies
// ST_HmiCommand to the plant. The HMI only ever sees these two structs.
// Commands that trigger an action act on the rising edge.
FUNCTION_BLOCK FB_HmiBridge
VAR_OUTPUT
    eModeRequest : E_OpMode := E_OpMode.eAutomatic;   // for MAIN's mode handler
END_VAR
VAR
    fbTeachStart   : R_TRIG;
    fbTeachConfirm : R_TRIG;
    fbResetFault   : R_TRIG;
END_VAR

METHOD PUBLIC Run
VAR_IN_OUT
    fbPlant  : FB_Hrl;
    fbEmu    : FB_MfrEmulator;
    stCmd    : ST_HmiCommand;
    stStat   : ST_HmiStatus;
END_VAR
VAR_INPUT
    eModeNow : E_OpMode;
END_VAR
VAR
    stAddr : ST_SlotAddr;
    i, nShown : INT;
    eJog : E_JogAxis;
END_VAR
// ---- HMI -> PLC
IF stCmd.bModeStop THEN            // stop wins if several are pressed
    eModeRequest := E_OpMode.eStop;
ELSIF stCmd.bModeManual THEN
    eModeRequest := E_OpMode.eManual;
ELSIF stCmd.bModeHoming THEN
    eModeRequest := E_OpMode.eHoming;
ELSIF stCmd.bModeAuto THEN
    eModeRequest := E_OpMode.eAutomatic;
END_IF
CASE stCmd.nJogAxis OF
    1: eJog := E_JogAxis.eHoist;
    2: eJog := E_JogAxis.eFork;
ELSE
    eJog := E_JogAxis.eTravel;
END_CASE
fbPlant.Jog(eJog, stCmd.bJogFwd, stCmd.bJogBwd);
fbPlant.bSafetyReset  := stCmd.bSafetyReset;
fbTeachStart(CLK := stCmd.bTeachStart);
IF fbTeachStart.Q THEN
    stAddr.nSide   := stCmd.nTeachSide;
    stAddr.nColumn := stCmd.nTeachColumn;
    stAddr.nLevel  := stCmd.nTeachLevel;
    fbPlant.fbTeach.Start(stAddr);
END_IF
fbTeachConfirm(CLK := stCmd.bTeachConfirm);
IF fbTeachConfirm.Q THEN
    fbPlant.fbTeach.Confirm();
END_IF
fbResetFault(CLK := stCmd.bResetFault);
IF fbResetFault.Q THEN
    fbPlant.fbSrm.ResetFault();
END_IF

// ---- PLC -> HMI
stStat.nMode         := TO_INT(eModeNow);
stStat.bSafetyOk     := fbPlant.bSafetyOk;
stStat.lrTravelPos   := fbPlant.fbSrm.TravelPos;
stStat.lrHoistPos    := fbPlant.fbSrm.HoistPos;
stStat.lrForkPos     := fbPlant.fbSrm.ForkActPos;
stStat.bBusy         := fbPlant.fbSrm.bBusy;
stStat.bFault        := fbPlant.fbSrm.bFault;
stStat.bJogBlocked   := fbPlant.fbSrm.bJogBlocked;
stStat.sLeOnFork     := fbPlant.fbSrm.sLeOnFork;
stStat.nJobsDone     := fbPlant.fbSrm.nJobsDone;
stStat.nStored       := fbEmu.nStored;
stStat.nRetrieved    := fbEmu.nRetrieved;
stStat.bMfrConnected := fbPlant.fbMfrTcp.bConnected;
stStat.nActiveFaults := fbPlant.fbDiag.nActive;
stStat.bTeachActive  := fbPlant.fbTeach.bActive;
stStat.nTaught       := fbPlant.fbTeach.nTaught;
stStat.bTeachRejected := fbPlant.fbTeach.bLastRejected;
stStat.sConfigError  := fbPlant.sConfigError;
stStat.sFault1 := ''; stStat.sFault2 := ''; stStat.sFault3 := ''; stStat.sFault4 := '';
nShown := 0;
FOR i := 1 TO 16 DO   // FB_Diag.cMaxFault
    IF fbPlant.fbDiag.aText[i] <> '' THEN
        nShown := nShown + 1;
        CASE nShown OF
            1: stStat.sFault1 := fbPlant.fbDiag.aText[i];
            2: stStat.sFault2 := fbPlant.fbDiag.aText[i];
            3: stStat.sFault3 := fbPlant.fbDiag.aText[i];
            4: stStat.sFault4 := fbPlant.fbDiag.aText[i];
        END_CASE
    END_IF
END_FOR
END_METHOD

END_FUNCTION_BLOCK

// ---- Test/PRG_TEST.TcPOU
// PRG_TEST - runs the unit tests with TcUnit. PlcTask calls it after MAIN; the
// suites build their own instances and never touch MAIN's plant. Results land
// in the Error List about a second after Run.
PROGRAM PRG_TEST
VAR
    fbRackTest      : FB_Rack_Test;
    fbAxisTest      : FB_Axis_Test;
    fbConveyorTest  : FB_ConveyorZone_Test;
    fbIPointTest    : FB_IPoint_Test;
    fbMfrTest       : FB_MfrInterface_Test;
    fbSrmTest       : FB_Srm_Test;
    fbTravelTimeTest: FB_TravelTime_Test;
    fbAxisNcTest    : FB_AxisNc_Test;
    fbConfigTest    : FB_HrlConfig_Test;
    fbCodecTest     : FB_TelegramCodec_Test;
    fbOperationTest : FB_Operation_Test;
    fbSafetyTest    : FB_SafetyInterface_Test;
END_VAR

TcUnit.RUN();

END_PROGRAM

// ---- Test/FB_Rack_Test.TcPOU
// Tests for FB_Rack: place geometry, teach-in, booking pallets in and out.
// Every test gets its own rack so they cannot see each other's pallets.
FUNCTION_BLOCK FB_Rack_Test EXTENDS TcUnit.FB_TestSuite
VAR
    fbRackGeo   : FB_Rack;
    fbRackTeach : FB_Rack;
    fbRackReject: FB_Rack;
    fbRackBook  : FB_Rack;
    fbRackTwice : FB_Rack;
    fbRackBad   : FB_Rack;
    fbRackFree  : FB_Rack;
END_VAR

Geometry_PlaceAndStation_FollowTheDrawing();
Teach_WithinTolerance_IsUsedAsTarget();
Teach_OutOfTolerance_IsRejected();
PutTake_BooksThePalletInAndOut();
Put_OnOccupiedPlace_IsRefused();
InvalidAddress_IsRejectedEverywhere();
FindFree_SkipsOccupiedPlaces();

METHOD PRIVATE Geometry_PlaceAndStation_FollowTheDrawing
VAR_INST
    bRan : BOOL;
END_VAR
VAR
    stPlace   : ST_SlotAddr := (nSide := 2, nColumn := 5, nLevel := 3);
    stStation : ST_SlotAddr := (nSide := 1, nColumn := 0, nLevel := 1);
END_VAR
TEST('Geometry_PlaceAndStation_FollowTheDrawing');
IF bRan THEN
    TEST_FINISHED();
    RETURN;
END_IF
bRan := TRUE;

AssertEquals_LREAL(Expected := 7.6, Actual := fbRackGeo.NominalX(stPlace), Delta := 1.0E-9, Message := 'column 5 = offset 2.0 + 4 x 1.4 m');
AssertEquals_LREAL(Expected := 3.1, Actual := fbRackGeo.NominalY(stPlace), Delta := 1.0E-9, Message := 'level 3 = offset 0.5 + 2 x 1.3 m');
AssertEquals_LREAL(Expected := 0.0, Actual := fbRackGeo.NominalX(stStation), Delta := 1.0E-9, Message := 'transfer station is the travel zero');
AssertTrue(Condition := fbRackGeo.IsStation(stStation), Message := 'column 0 / level 1 / side 1 is the station');

TEST_FINISHED();
END_METHOD

METHOD PRIVATE Teach_WithinTolerance_IsUsedAsTarget
VAR_INST
    bRan : BOOL;
END_VAR
VAR
    stPlace : ST_SlotAddr := (nSide := 1, nColumn := 3, nLevel := 2);
    lrX, lrY : LREAL;
END_VAR
TEST('Teach_WithinTolerance_IsUsedAsTarget');
IF bRan THEN
    TEST_FINISHED();
    RETURN;
END_IF
bRan := TRUE;

lrX := fbRackTeach.NominalX(stPlace) + 0.012;
lrY := fbRackTeach.NominalY(stPlace) - 0.008;
AssertTrue(Condition := fbRackTeach.Teach(stPlace, lrX, lrY), Message := '12 mm / 8 mm off the drawing must be accepted');
AssertEquals_LREAL(Expected := lrX, Actual := fbRackTeach.TargetX(stPlace), Delta := 1.0E-9, Message := 'RBG must drive to the taught travel position');
AssertEquals_LREAL(Expected := lrY, Actual := fbRackTeach.TargetY(stPlace), Delta := 1.0E-9, Message := 'RBG must drive to the taught hoist position');

TEST_FINISHED();
END_METHOD

